REGION Network 43: Barcode - System 3
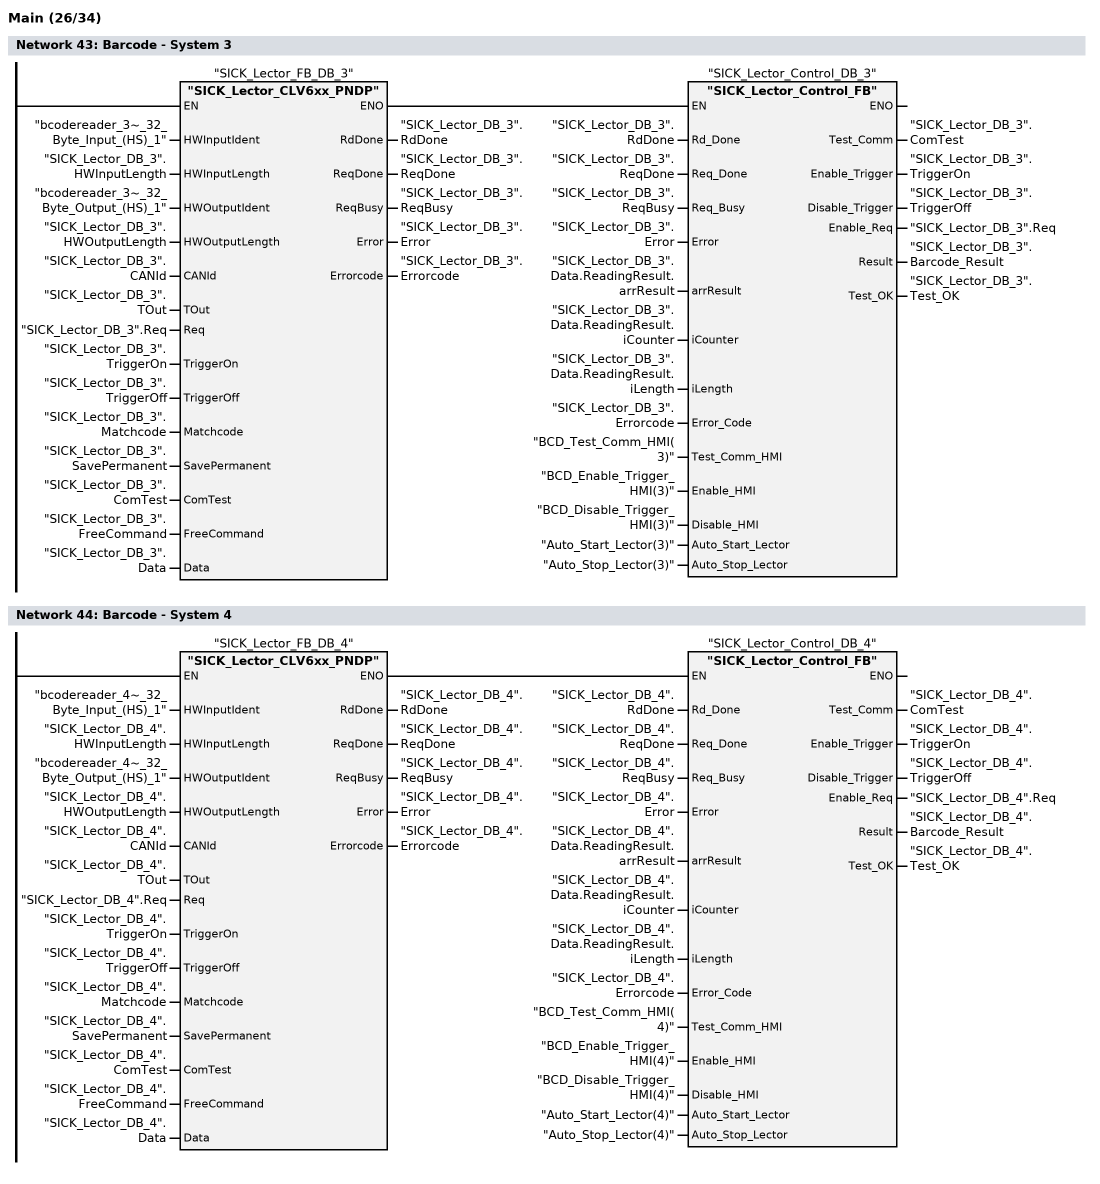
   RUNG wire#powerrail
      "SICK_Lector_FB_DB_3"(HWInputIdent := "bcodereader_3~_32_Byte_Input_(HS)_1", HWInputLength := "SICK_Lector_DB_3".HWInputLength, HWOutputIdent := "bcodereader_3~_32_Byte_Output_(HS)_1", HWOutputLength := "SICK_Lector_DB_3".HWOutputLength, CANId := "SICK_Lector_DB_3".CANId, TOut := "SICK_Lector_DB_3".TOut, Req := "SICK_Lector_DB_3".Req, TriggerOn := "SICK_Lector_DB_3".TriggerOn, TriggerOff := "SICK_Lector_DB_3".TriggerOff, Matchcode := "SICK_Lector_DB_3".Matchcode, SavePermanent := "SICK_Lector_DB_3".SavePermanent, ComTest := "SICK_Lector_DB_3".ComTest, FreeCommand := "SICK_Lector_DB_3".FreeCommand, Data := "SICK_Lector_DB_3".Data, RdDone => "SICK_Lector_DB_3".RdDone, ReqDone => "SICK_Lector_DB_3".ReqDone, ReqBusy => "SICK_Lector_DB_3".ReqBusy, Error => "SICK_Lector_DB_3".Error, Errorcode => "SICK_Lector_DB_3".Errorcode)
      "SICK_Lector_Control_DB_3"(Rd_Done := "SICK_Lector_DB_3".RdDone, Req_Done := "SICK_Lector_DB_3".ReqDone, Req_Busy := "SICK_Lector_DB_3".ReqBusy, Error := "SICK_Lector_DB_3".Error, arrResult := "SICK_Lector_DB_3".Data.ReadingResult.arrResult, iCounter := "SICK_Lector_DB_3".Data.ReadingResult.iCounter, iLength := "SICK_Lector_DB_3".Data.ReadingResult.iLength, Error_Code := "SICK_Lector_DB_3".Errorcode, Test_Comm_HMI := "BCD_Test_Comm_HMI(3)", Enable_HMI := "BCD_Enable_Trigger_HMI(3)", Disable_HMI := "BCD_Disable_Trigger_HMI(3)", Auto_Start_Lector := "Auto_Start_Lector(3)", Auto_Stop_Lector := "Auto_Stop_Lector(3)", Test_Comm => "SICK_Lector_DB_3".ComTest, Enable_Trigger => "SICK_Lector_DB_3".TriggerOn, Disable_Trigger => "SICK_Lector_DB_3".TriggerOff, Enable_Req => "SICK_Lector_DB_3".Req, Result => "SICK_Lector_DB_3".Barcode_Result, Test_OK => "SICK_Lector_DB_3".Test_OK)
   END_RUNG
   // the same network as SCL:
   "SICK_Lector_FB_DB_3"(HWInputIdent := "bcodereader_3~_32_Byte_Input_(HS)_1",   // "SICK_Lector_CLV6xx_PNDP"
                         HWInputLength := "SICK_Lector_DB_3".HWInputLength,
                         HWOutputIdent := "bcodereader_3~_32_Byte_Output_(HS)_1",
                         HWOutputLength := "SICK_Lector_DB_3".HWOutputLength,
                         CANId := "SICK_Lector_DB_3".CANId,
                         TOut := "SICK_Lector_DB_3".TOut,
                         Req := "SICK_Lector_DB_3".Req,
                         TriggerOn := "SICK_Lector_DB_3".TriggerOn,
                         TriggerOff := "SICK_Lector_DB_3".TriggerOff,
                         Matchcode := "SICK_Lector_DB_3".Matchcode,
                         SavePermanent := "SICK_Lector_DB_3".SavePermanent,
                         ComTest := "SICK_Lector_DB_3".ComTest,
                         FreeCommand := "SICK_Lector_DB_3".FreeCommand,
                         Data := "SICK_Lector_DB_3".Data,
                         RdDone => "SICK_Lector_DB_3".RdDone,
                         ReqDone => "SICK_Lector_DB_3".ReqDone,
                         ReqBusy => "SICK_Lector_DB_3".ReqBusy,
                         Error => "SICK_Lector_DB_3".Error,
                         Errorcode => "SICK_Lector_DB_3".Errorcode,
                         ENO => #_w1);
   IF #_w1 THEN
       "SICK_Lector_Control_DB_3"(Rd_Done := "SICK_Lector_DB_3".RdDone,   // "SICK_Lector_Control_FB"
                               Req_Done := "SICK_Lector_DB_3".ReqDone,
                               Req_Busy := "SICK_Lector_DB_3".ReqBusy,
                               Error := "SICK_Lector_DB_3".Error,
                               arrResult := "SICK_Lector_DB_3".Data.ReadingResult.arrResult,
                               iCounter := "SICK_Lector_DB_3".Data.ReadingResult.iCounter,
                               iLength := "SICK_Lector_DB_3".Data.ReadingResult.iLength,
                               Error_Code := "SICK_Lector_DB_3".Errorcode,
                               Test_Comm_HMI := "BCD_Test_Comm_HMI(3)",
                               Enable_HMI := "BCD_Enable_Trigger_HMI(3)",
                               Disable_HMI := "BCD_Disable_Trigger_HMI(3)",
                               Auto_Start_Lector := "Auto_Start_Lector(3)",
                               Auto_Stop_Lector := "Auto_Stop_Lector(3)",
                               Test_Comm => "SICK_Lector_DB_3".ComTest,
                               Enable_Trigger => "SICK_Lector_DB_3".TriggerOn,
                               Disable_Trigger => "SICK_Lector_DB_3".TriggerOff,
                               Enable_Req => "SICK_Lector_DB_3".Req,
                               Result => "SICK_Lector_DB_3".Barcode_Result,
                               Test_OK => "SICK_Lector_DB_3".Test_OK);
   END_IF;
END_REGION

REGION Network 44: Barcode - System 4
   RUNG wire#powerrail
      "SICK_Lector_FB_DB_4"(HWInputIdent := "bcodereader_4~_32_Byte_Input_(HS)_1", HWInputLength := "SICK_Lector_DB_4".HWInputLength, HWOutputIdent := "bcodereader_4~_32_Byte_Output_(HS)_1", HWOutputLength := "SICK_Lector_DB_4".HWOutputLength, CANId := "SICK_Lector_DB_4".CANId, TOut := "SICK_Lector_DB_4".TOut, Req := "SICK_Lector_DB_4".Req, TriggerOn := "SICK_Lector_DB_4".TriggerOn, TriggerOff := "SICK_Lector_DB_4".TriggerOff, Matchcode := "SICK_Lector_DB_4".Matchcode, SavePermanent := "SICK_Lector_DB_4".SavePermanent, ComTest := "SICK_Lector_DB_4".ComTest, FreeCommand := "SICK_Lector_DB_4".FreeCommand, Data := "SICK_Lector_DB_4".Data, RdDone => "SICK_Lector_DB_4".RdDone, ReqDone => "SICK_Lector_DB_4".ReqDone, ReqBusy => "SICK_Lector_DB_4".ReqBusy, Error => "SICK_Lector_DB_4".Error, Errorcode => "SICK_Lector_DB_4".Errorcode)
      "SICK_Lector_Control_DB_4"(Rd_Done := "SICK_Lector_DB_4".RdDone, Req_Done := "SICK_Lector_DB_4".ReqDone, Req_Busy := "SICK_Lector_DB_4".ReqBusy, Error := "SICK_Lector_DB_4".Error, arrResult := "SICK_Lector_DB_4".Data.ReadingResult.arrResult, iCounter := "SICK_Lector_DB_4".Data.ReadingResult.iCounter, iLength := "SICK_Lector_DB_4".Data.ReadingResult.iLength, Error_Code := "SICK_Lector_DB_4".Errorcode, Test_Comm_HMI := "BCD_Test_Comm_HMI(4)", Enable_HMI := "BCD_Enable_Trigger_HMI(4)", Disable_HMI := "BCD_Disable_Trigger_HMI(4)", Auto_Start_Lector := "Auto_Start_Lector(4)", Auto_Stop_Lector := "Auto_Stop_Lector(4)", Test_Comm => "SICK_Lector_DB_4".ComTest, Enable_Trigger => "SICK_Lector_DB_4".TriggerOn, Disable_Trigger => "SICK_Lector_DB_4".TriggerOff, Enable_Req => "SICK_Lector_DB_4".Req, Result => "SICK_Lector_DB_4".Barcode_Result, Test_OK => "SICK_Lector_DB_4".Test_OK)
   END_RUNG
   // the same network as SCL:
   "SICK_Lector_FB_DB_4"(HWInputIdent := "bcodereader_4~_32_Byte_Input_(HS)_1",   // "SICK_Lector_CLV6xx_PNDP"
                         HWInputLength := "SICK_Lector_DB_4".HWInputLength,
                         HWOutputIdent := "bcodereader_4~_32_Byte_Output_(HS)_1",
                         HWOutputLength := "SICK_Lector_DB_4".HWOutputLength,
                         CANId := "SICK_Lector_DB_4".CANId,
                         TOut := "SICK_Lector_DB_4".TOut,
                         Req := "SICK_Lector_DB_4".Req,
                         TriggerOn := "SICK_Lector_DB_4".TriggerOn,
                         TriggerOff := "SICK_Lector_DB_4".TriggerOff,
                         Matchcode := "SICK_Lector_DB_4".Matchcode,
                         SavePermanent := "SICK_Lector_DB_4".SavePermanent,
                         ComTest := "SICK_Lector_DB_4".ComTest,
                         FreeCommand := "SICK_Lector_DB_4".FreeCommand,
                         Data := "SICK_Lector_DB_4".Data,
                         RdDone => "SICK_Lector_DB_4".RdDone,
                         ReqDone => "SICK_Lector_DB_4".ReqDone,
                         ReqBusy => "SICK_Lector_DB_4".ReqBusy,
                         Error => "SICK_Lector_DB_4".Error,
                         Errorcode => "SICK_Lector_DB_4".Errorcode,
                         ENO => #_w1);
   IF #_w1 THEN
       "SICK_Lector_Control_DB_4"(Rd_Done := "SICK_Lector_DB_4".RdDone,   // "SICK_Lector_Control_FB"
                               Req_Done := "SICK_Lector_DB_4".ReqDone,
                               Req_Busy := "SICK_Lector_DB_4".ReqBusy,
                               Error := "SICK_Lector_DB_4".Error,
                               arrResult := "SICK_Lector_DB_4".Data.ReadingResult.arrResult,
                               iCounter := "SICK_Lector_DB_4".Data.ReadingResult.iCounter,
                               iLength := "SICK_Lector_DB_4".Data.ReadingResult.iLength,
                               Error_Code := "SICK_Lector_DB_4".Errorcode,
                               Test_Comm_HMI := "BCD_Test_Comm_HMI(4)",
                               Enable_HMI := "BCD_Enable_Trigger_HMI(4)",
                               Disable_HMI := "BCD_Disable_Trigger_HMI(4)",
                               Auto_Start_Lector := "Auto_Start_Lector(4)",
                               Auto_Stop_Lector := "Auto_Stop_Lector(4)",
                               Test_Comm => "SICK_Lector_DB_4".ComTest,
                               Enable_Trigger => "SICK_Lector_DB_4".TriggerOn,
                               Disable_Trigger => "SICK_Lector_DB_4".TriggerOff,
                               Enable_Req => "SICK_Lector_DB_4".Req,
                               Result => "SICK_Lector_DB_4".Barcode_Result,
                               Test_OK => "SICK_Lector_DB_4".Test_OK);
   END_IF;
END_REGION

REGION Network 45: Barcode - System 5
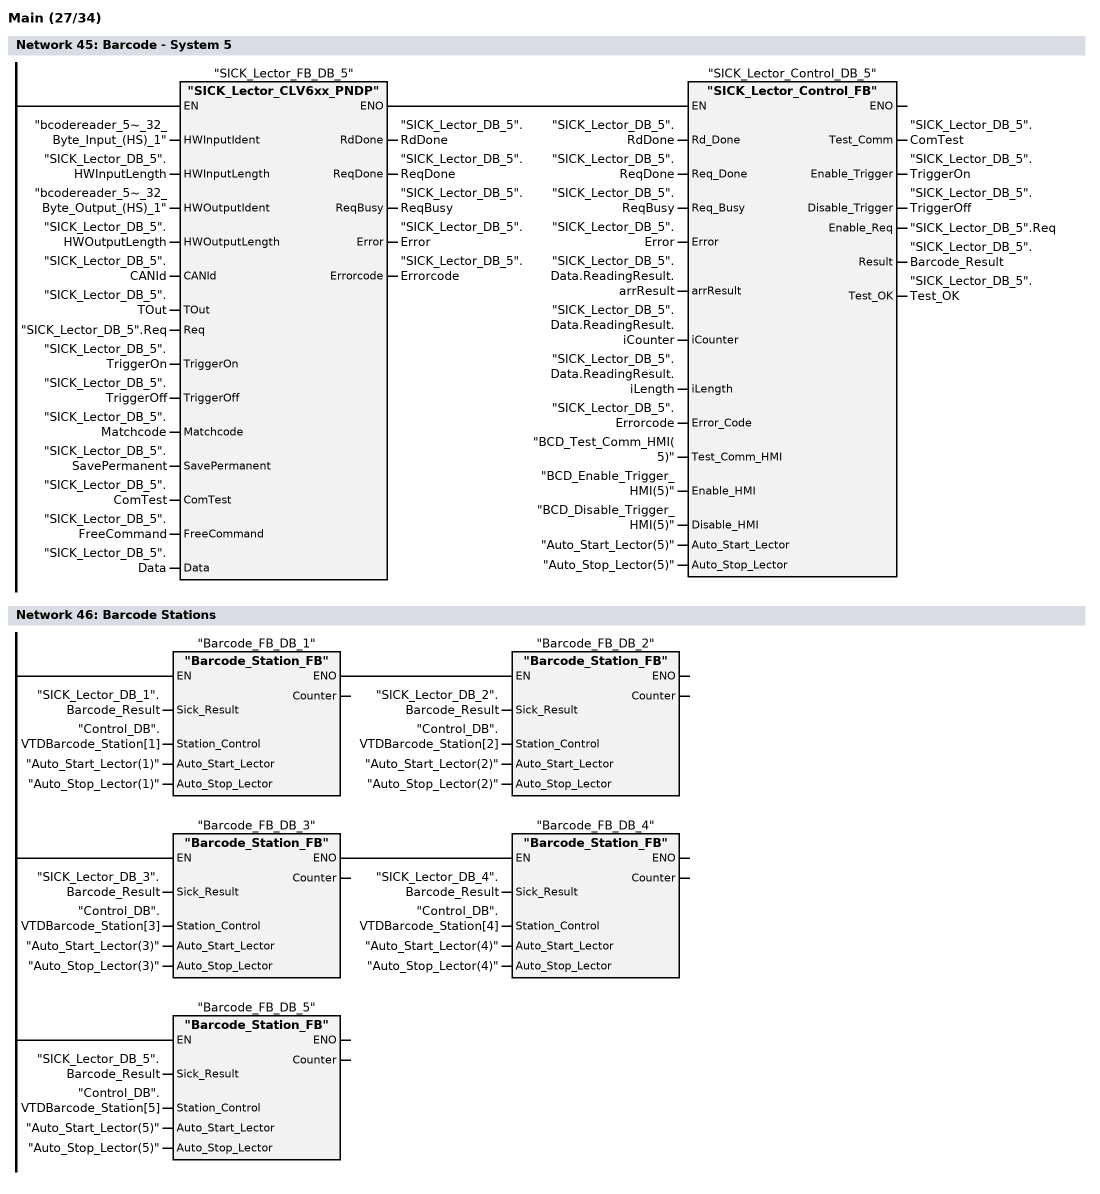
   RUNG wire#powerrail
      "SICK_Lector_FB_DB_5"(HWInputIdent := "bcodereader_5~_32_Byte_Input_(HS)_1", HWInputLength := "SICK_Lector_DB_5".HWInputLength, HWOutputIdent := "bcodereader_5~_32_Byte_Output_(HS)_1", HWOutputLength := "SICK_Lector_DB_5".HWOutputLength, CANId := "SICK_Lector_DB_5".CANId, TOut := "SICK_Lector_DB_5".TOut, Req := "SICK_Lector_DB_5".Req, TriggerOn := "SICK_Lector_DB_5".TriggerOn, TriggerOff := "SICK_Lector_DB_5".TriggerOff, Matchcode := "SICK_Lector_DB_5".Matchcode, SavePermanent := "SICK_Lector_DB_5".SavePermanent, ComTest := "SICK_Lector_DB_5".ComTest, FreeCommand := "SICK_Lector_DB_5".FreeCommand, Data := "SICK_Lector_DB_5".Data, RdDone => "SICK_Lector_DB_5".RdDone, ReqDone => "SICK_Lector_DB_5".ReqDone, ReqBusy => "SICK_Lector_DB_5".ReqBusy, Error => "SICK_Lector_DB_5".Error, Errorcode => "SICK_Lector_DB_5".Errorcode)
      "SICK_Lector_Control_DB_5"(Rd_Done := "SICK_Lector_DB_5".RdDone, Req_Done := "SICK_Lector_DB_5".ReqDone, Req_Busy := "SICK_Lector_DB_5".ReqBusy, Error := "SICK_Lector_DB_5".Error, arrResult := "SICK_Lector_DB_5".Data.ReadingResult.arrResult, iCounter := "SICK_Lector_DB_5".Data.ReadingResult.iCounter, iLength := "SICK_Lector_DB_5".Data.ReadingResult.iLength, Error_Code := "SICK_Lector_DB_5".Errorcode, Test_Comm_HMI := "BCD_Test_Comm_HMI(5)", Enable_HMI := "BCD_Enable_Trigger_HMI(5)", Disable_HMI := "BCD_Disable_Trigger_HMI(5)", Auto_Start_Lector := "Auto_Start_Lector(5)", Auto_Stop_Lector := "Auto_Stop_Lector(5)", Test_Comm => "SICK_Lector_DB_5".ComTest, Enable_Trigger => "SICK_Lector_DB_5".TriggerOn, Disable_Trigger => "SICK_Lector_DB_5".TriggerOff, Enable_Req => "SICK_Lector_DB_5".Req, Result => "SICK_Lector_DB_5".Barcode_Result, Test_OK => "SICK_Lector_DB_5".Test_OK)
   END_RUNG
   // the same network as SCL:
   "SICK_Lector_FB_DB_5"(HWInputIdent := "bcodereader_5~_32_Byte_Input_(HS)_1",   // "SICK_Lector_CLV6xx_PNDP"
                         HWInputLength := "SICK_Lector_DB_5".HWInputLength,
                         HWOutputIdent := "bcodereader_5~_32_Byte_Output_(HS)_1",
                         HWOutputLength := "SICK_Lector_DB_5".HWOutputLength,
                         CANId := "SICK_Lector_DB_5".CANId,
                         TOut := "SICK_Lector_DB_5".TOut,
                         Req := "SICK_Lector_DB_5".Req,
                         TriggerOn := "SICK_Lector_DB_5".TriggerOn,
                         TriggerOff := "SICK_Lector_DB_5".TriggerOff,
                         Matchcode := "SICK_Lector_DB_5".Matchcode,
                         SavePermanent := "SICK_Lector_DB_5".SavePermanent,
                         ComTest := "SICK_Lector_DB_5".ComTest,
                         FreeCommand := "SICK_Lector_DB_5".FreeCommand,
                         Data := "SICK_Lector_DB_5".Data,
                         RdDone => "SICK_Lector_DB_5".RdDone,
                         ReqDone => "SICK_Lector_DB_5".ReqDone,
                         ReqBusy => "SICK_Lector_DB_5".ReqBusy,
                         Error => "SICK_Lector_DB_5".Error,
                         Errorcode => "SICK_Lector_DB_5".Errorcode,
                         ENO => #_w1);
   IF #_w1 THEN
       "SICK_Lector_Control_DB_5"(Rd_Done := "SICK_Lector_DB_5".RdDone,   // "SICK_Lector_Control_FB"
                               Req_Done := "SICK_Lector_DB_5".ReqDone,
                               Req_Busy := "SICK_Lector_DB_5".ReqBusy,
                               Error := "SICK_Lector_DB_5".Error,
                               arrResult := "SICK_Lector_DB_5".Data.ReadingResult.arrResult,
                               iCounter := "SICK_Lector_DB_5".Data.ReadingResult.iCounter,
                               iLength := "SICK_Lector_DB_5".Data.ReadingResult.iLength,
                               Error_Code := "SICK_Lector_DB_5".Errorcode,
                               Test_Comm_HMI := "BCD_Test_Comm_HMI(5)",
                               Enable_HMI := "BCD_Enable_Trigger_HMI(5)",
                               Disable_HMI := "BCD_Disable_Trigger_HMI(5)",
                               Auto_Start_Lector := "Auto_Start_Lector(5)",
                               Auto_Stop_Lector := "Auto_Stop_Lector(5)",
                               Test_Comm => "SICK_Lector_DB_5".ComTest,
                               Enable_Trigger => "SICK_Lector_DB_5".TriggerOn,
                               Disable_Trigger => "SICK_Lector_DB_5".TriggerOff,
                               Enable_Req => "SICK_Lector_DB_5".Req,
                               Result => "SICK_Lector_DB_5".Barcode_Result,
                               Test_OK => "SICK_Lector_DB_5".Test_OK);
   END_IF;
END_REGION

REGION Network 46: Barcode Stations
   RUNG wire#powerrail
      "Barcode_FB_DB_1"(Sick_Result := "SICK_Lector_DB_1".Barcode_Result, Station_Control := "Control_DB".VTDBarcode_Station[1], Auto_Start_Lector := "Auto_Start_Lector(1)", Auto_Stop_Lector := "Auto_Stop_Lector(1)", "Counter" =>)
      "Barcode_FB_DB_2"(Sick_Result := "SICK_Lector_DB_2".Barcode_Result, Station_Control := "Control_DB".VTDBarcode_Station[2], Auto_Start_Lector := "Auto_Start_Lector(2)", Auto_Stop_Lector := "Auto_Stop_Lector(2)", "Counter" =>)
   END_RUNG
   RUNG wire#powerrail
      "Barcode_FB_DB_3"(Sick_Result := "SICK_Lector_DB_3".Barcode_Result, Station_Control := "Control_DB".VTDBarcode_Station[3], Auto_Start_Lector := "Auto_Start_Lector(3)", Auto_Stop_Lector := "Auto_Stop_Lector(3)", "Counter" =>)
      "Barcode_FB_DB_4"(Sick_Result := "SICK_Lector_DB_4".Barcode_Result, Station_Control := "Control_DB".VTDBarcode_Station[4], Auto_Start_Lector := "Auto_Start_Lector(4)", Auto_Stop_Lector := "Auto_Stop_Lector(4)", "Counter" =>)
   END_RUNG
   RUNG wire#powerrail
      "Barcode_FB_DB_5"(Sick_Result := "SICK_Lector_DB_5".Barcode_Result, Station_Control := "Control_DB".VTDBarcode_Station[5], Auto_Start_Lector := "Auto_Start_Lector(5)", Auto_Stop_Lector := "Auto_Stop_Lector(5)", "Counter" =>)
   END_RUNG
   // the same network as SCL:
   "Barcode_FB_DB_1"(Sick_Result := "SICK_Lector_DB_1".Barcode_Result,   // "Barcode_Station_FB"
                     Station_Control := "Control_DB".VTDBarcode_Station[1],
                     Auto_Start_Lector := "Auto_Start_Lector(1)",
                     Auto_Stop_Lector := "Auto_Stop_Lector(1)",
                     ENO => #_w1);
   IF #_w1 THEN
       "Barcode_FB_DB_2"(Sick_Result := "SICK_Lector_DB_2".Barcode_Result,   // "Barcode_Station_FB"
                         Station_Control := "Control_DB".VTDBarcode_Station[2],
                         Auto_Start_Lector := "Auto_Start_Lector(2)",
                         Auto_Stop_Lector := "Auto_Stop_Lector(2)");
   END_IF;
   "Barcode_FB_DB_3"(Sick_Result := "SICK_Lector_DB_3".Barcode_Result,   // "Barcode_Station_FB"
                     Station_Control := "Control_DB".VTDBarcode_Station[3],
                     Auto_Start_Lector := "Auto_Start_Lector(3)",
                     Auto_Stop_Lector := "Auto_Stop_Lector(3)",
                     ENO => #_w2);
   IF #_w2 THEN
       "Barcode_FB_DB_4"(Sick_Result := "SICK_Lector_DB_4".Barcode_Result,   // "Barcode_Station_FB"
                         Station_Control := "Control_DB".VTDBarcode_Station[4],
                         Auto_Start_Lector := "Auto_Start_Lector(4)",
                         Auto_Stop_Lector := "Auto_Stop_Lector(4)");
   END_IF;
   "Barcode_FB_DB_5"(Sick_Result := "SICK_Lector_DB_5".Barcode_Result,   // "Barcode_Station_FB"
                     Station_Control := "Control_DB".VTDBarcode_Station[5],
                     Auto_Start_Lector := "Auto_Start_Lector(5)",
                     Auto_Stop_Lector := "Auto_Stop_Lector(5)");
END_REGION

REGION Network 47: Stack Lights
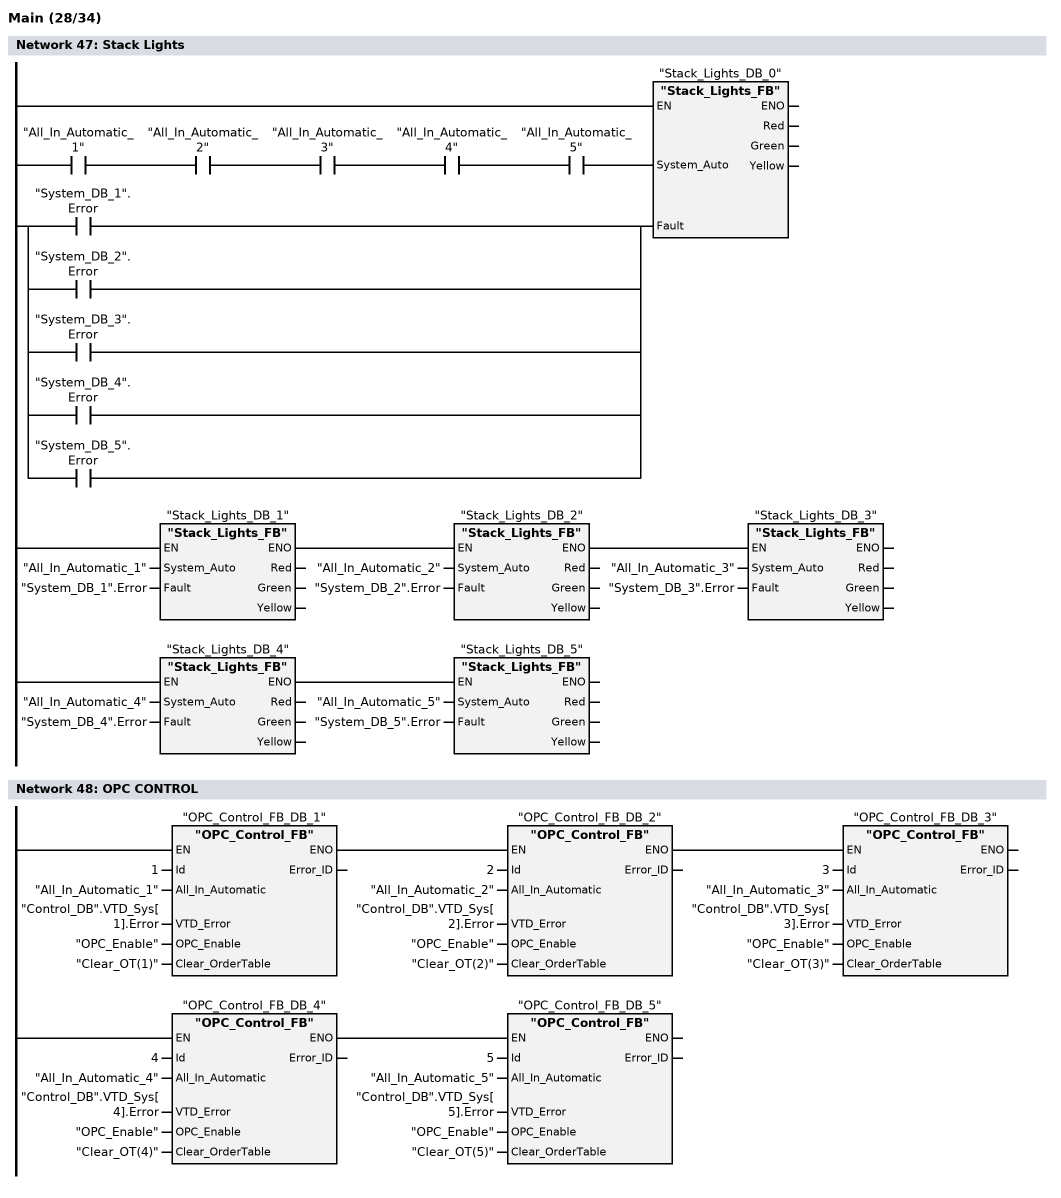
   RUNG wire#powerrail
      "Stack_Lights_DB_0"(System_Auto := wire#w1, Fault := wire#w2, Red =>, Green =>, Yellow =>)
   END_RUNG
   RUNG wire#powerrail
      Contact( "All_In_Automatic_1" )
      Contact( "All_In_Automatic_2" )
      Contact( "All_In_Automatic_3" )
      Contact( "All_In_Automatic_4" )
      Contact( "All_In_Automatic_5" )
   END_RUNG wire#w1
   RUNG wire#powerrail
      Contact( "System_DB_1".Error )
   END_RUNG wire#w2
   RUNG wire#powerrail
      Contact( "System_DB_2".Error )
   END_RUNG wire#w2
   RUNG wire#powerrail
      Contact( "System_DB_3".Error )
   END_RUNG wire#w2
   RUNG wire#powerrail
      Contact( "System_DB_4".Error )
   END_RUNG wire#w2
   RUNG wire#powerrail
      Contact( "System_DB_5".Error )
   END_RUNG wire#w2
   RUNG wire#powerrail
      "Stack_Lights_DB_1"(System_Auto := "All_In_Automatic_1", Fault := "System_DB_1".Error, Red =>, Green =>, Yellow =>)
      "Stack_Lights_DB_2"(System_Auto := "All_In_Automatic_2", Fault := "System_DB_2".Error, Red =>, Green =>, Yellow =>)
      "Stack_Lights_DB_3"(System_Auto := "All_In_Automatic_3", Fault := "System_DB_3".Error, Red =>, Green =>, Yellow =>)
   END_RUNG
   RUNG wire#powerrail
      "Stack_Lights_DB_4"(System_Auto := "All_In_Automatic_4", Fault := "System_DB_4".Error, Red =>, Green =>, Yellow =>)
      "Stack_Lights_DB_5"(System_Auto := "All_In_Automatic_5", Fault := "System_DB_5".Error, Red =>, Green =>, Yellow =>)
   END_RUNG
   // the same network as SCL:
   "Stack_Lights_DB_0"(System_Auto := "All_In_Automatic_1" AND "All_In_Automatic_2" AND "All_In_Automatic_3" AND "All_In_Automatic_4" AND "All_In_Automatic_5",   // "Stack_Lights_FB"
                       Fault := "System_DB_1".Error OR "System_DB_2".Error OR "System_DB_3".Error OR "System_DB_4".Error OR "System_DB_5".Error);
   "Stack_Lights_DB_1"(System_Auto := "All_In_Automatic_1", Fault := "System_DB_1".Error, ENO => #_w1);   // "Stack_Lights_FB"
   "Stack_Lights_DB_2"(EN := #_w1,   // "Stack_Lights_FB"
                       System_Auto := "All_In_Automatic_2",
                       Fault := "System_DB_2".Error,
                       ENO => #_w2);
   IF #_w2 THEN
       "Stack_Lights_DB_3"(System_Auto := "All_In_Automatic_3", Fault := "System_DB_3".Error);   // "Stack_Lights_FB"
   END_IF;
   "Stack_Lights_DB_4"(System_Auto := "All_In_Automatic_4", Fault := "System_DB_4".Error, ENO => #_w3);   // "Stack_Lights_FB"
   IF #_w3 THEN
       "Stack_Lights_DB_5"(System_Auto := "All_In_Automatic_5", Fault := "System_DB_5".Error);   // "Stack_Lights_FB"
   END_IF;
END_REGION

REGION Network 48: OPC CONTROL
   RUNG wire#powerrail
      "OPC_Control_FB_DB_1"(Id := 1, All_In_Automatic := "All_In_Automatic_1", VTD_Error := "Control_DB".VTD_Sys[1].Error, OPC_Enable := "OPC_Enable", Clear_OrderTable := "Clear_OT(1)", Error_ID =>)
      "OPC_Control_FB_DB_2"(Id := 2, All_In_Automatic := "All_In_Automatic_2", VTD_Error := "Control_DB".VTD_Sys[2].Error, OPC_Enable := "OPC_Enable", Clear_OrderTable := "Clear_OT(2)", Error_ID =>)
      "OPC_Control_FB_DB_3"(Id := 3, All_In_Automatic := "All_In_Automatic_3", VTD_Error := "Control_DB".VTD_Sys[3].Error, OPC_Enable := "OPC_Enable", Clear_OrderTable := "Clear_OT(3)", Error_ID =>)
   END_RUNG
   RUNG wire#powerrail
      "OPC_Control_FB_DB_4"(Id := 4, All_In_Automatic := "All_In_Automatic_4", VTD_Error := "Control_DB".VTD_Sys[4].Error, OPC_Enable := "OPC_Enable", Clear_OrderTable := "Clear_OT(4)", Error_ID =>)
      "OPC_Control_FB_DB_5"(Id := 5, All_In_Automatic := "All_In_Automatic_5", VTD_Error := "Control_DB".VTD_Sys[5].Error, OPC_Enable := "OPC_Enable", Clear_OrderTable := "Clear_OT(5)", Error_ID =>)
   END_RUNG
   // the same network as SCL:
   "OPC_Control_FB_DB_1"(Id := 1,   // "OPC_Control_FB"
                         All_In_Automatic := "All_In_Automatic_1",
                         VTD_Error := "Control_DB".VTD_Sys[1].Error,
                         OPC_Enable := "OPC_Enable",
                         Clear_OrderTable := "Clear_OT(1)",
                         ENO => #_w1);
   "OPC_Control_FB_DB_2"(EN := #_w1,   // "OPC_Control_FB"
                         Id := 2,
                         All_In_Automatic := "All_In_Automatic_2",
                         VTD_Error := "Control_DB".VTD_Sys[2].Error,
                         OPC_Enable := "OPC_Enable",
                         Clear_OrderTable := "Clear_OT(2)",
                         ENO => #_w2);
   IF #_w2 THEN
       "OPC_Control_FB_DB_3"(Id := 3,   // "OPC_Control_FB"
                             All_In_Automatic := "All_In_Automatic_3",
                             VTD_Error := "Control_DB".VTD_Sys[3].Error,
                             OPC_Enable := "OPC_Enable",
                             Clear_OrderTable := "Clear_OT(3)");
   END_IF;
   "OPC_Control_FB_DB_4"(Id := 4,   // "OPC_Control_FB"
                         All_In_Automatic := "All_In_Automatic_4",
                         VTD_Error := "Control_DB".VTD_Sys[4].Error,
                         OPC_Enable := "OPC_Enable",
                         Clear_OrderTable := "Clear_OT(4)",
                         ENO => #_w3);
   IF #_w3 THEN
       "OPC_Control_FB_DB_5"(Id := 5,   // "OPC_Control_FB"
                             All_In_Automatic := "All_In_Automatic_5",
                             VTD_Error := "Control_DB".VTD_Sys[5].Error,
                             OPC_Enable := "OPC_Enable",
                             Clear_OrderTable := "Clear_OT(5)");
   END_IF;
END_REGION

REGION Network 49: Shuttle TCPs
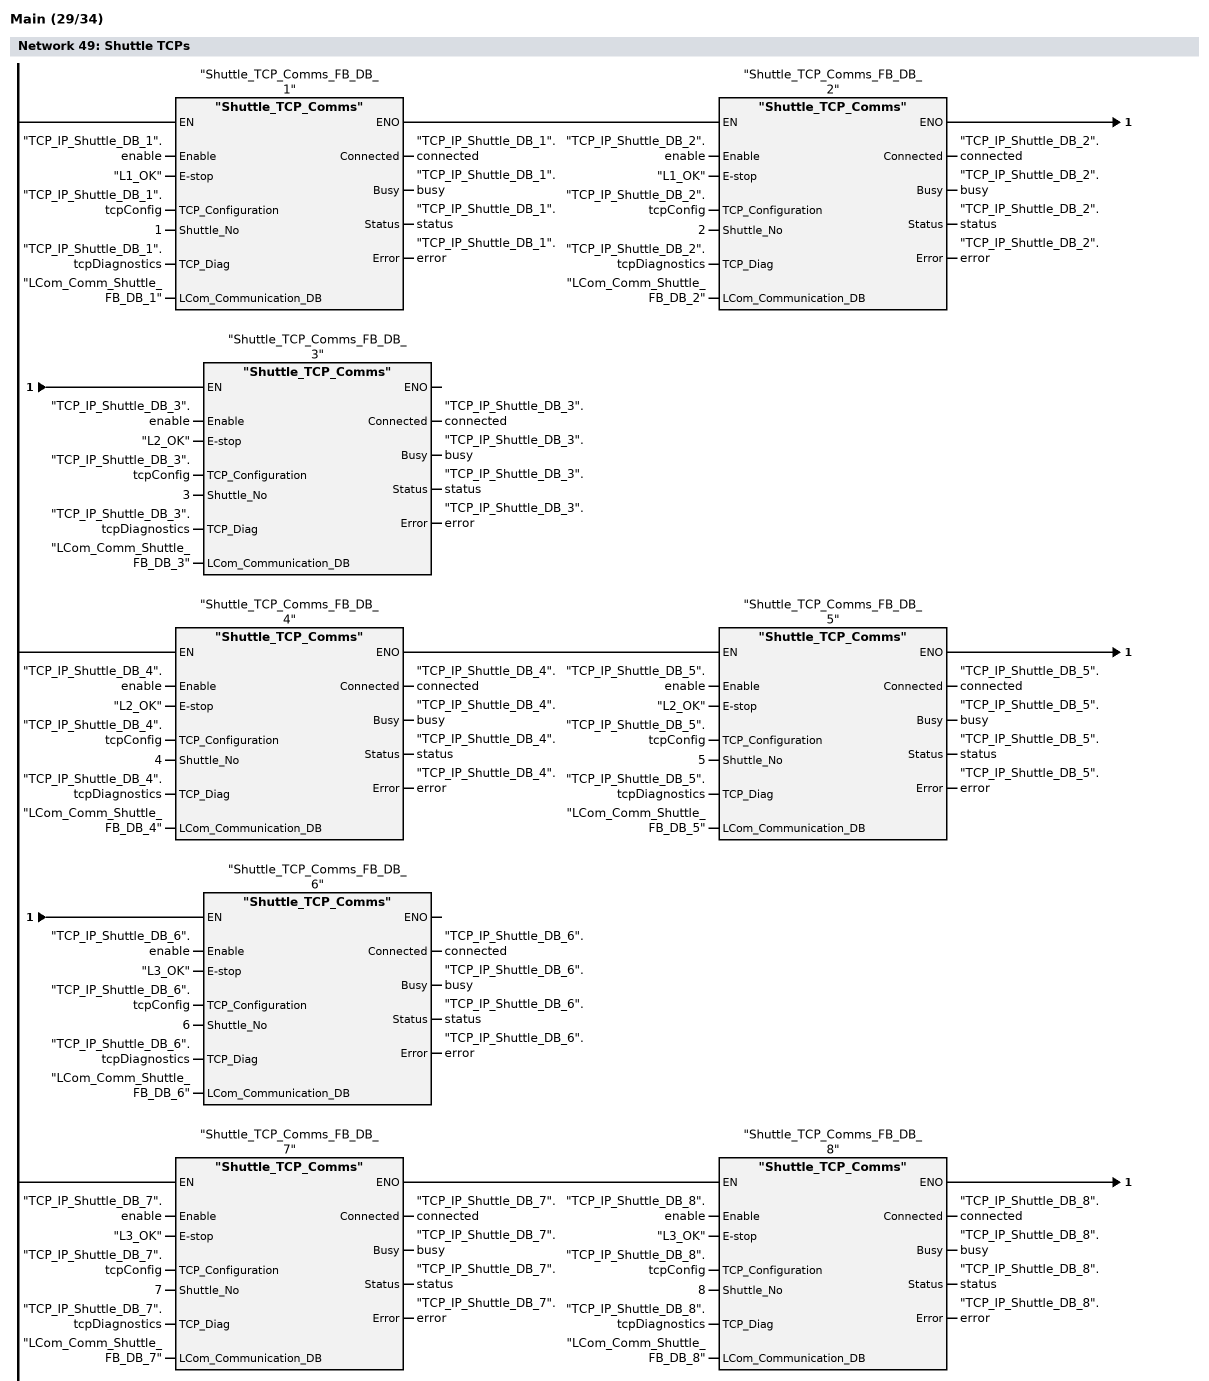
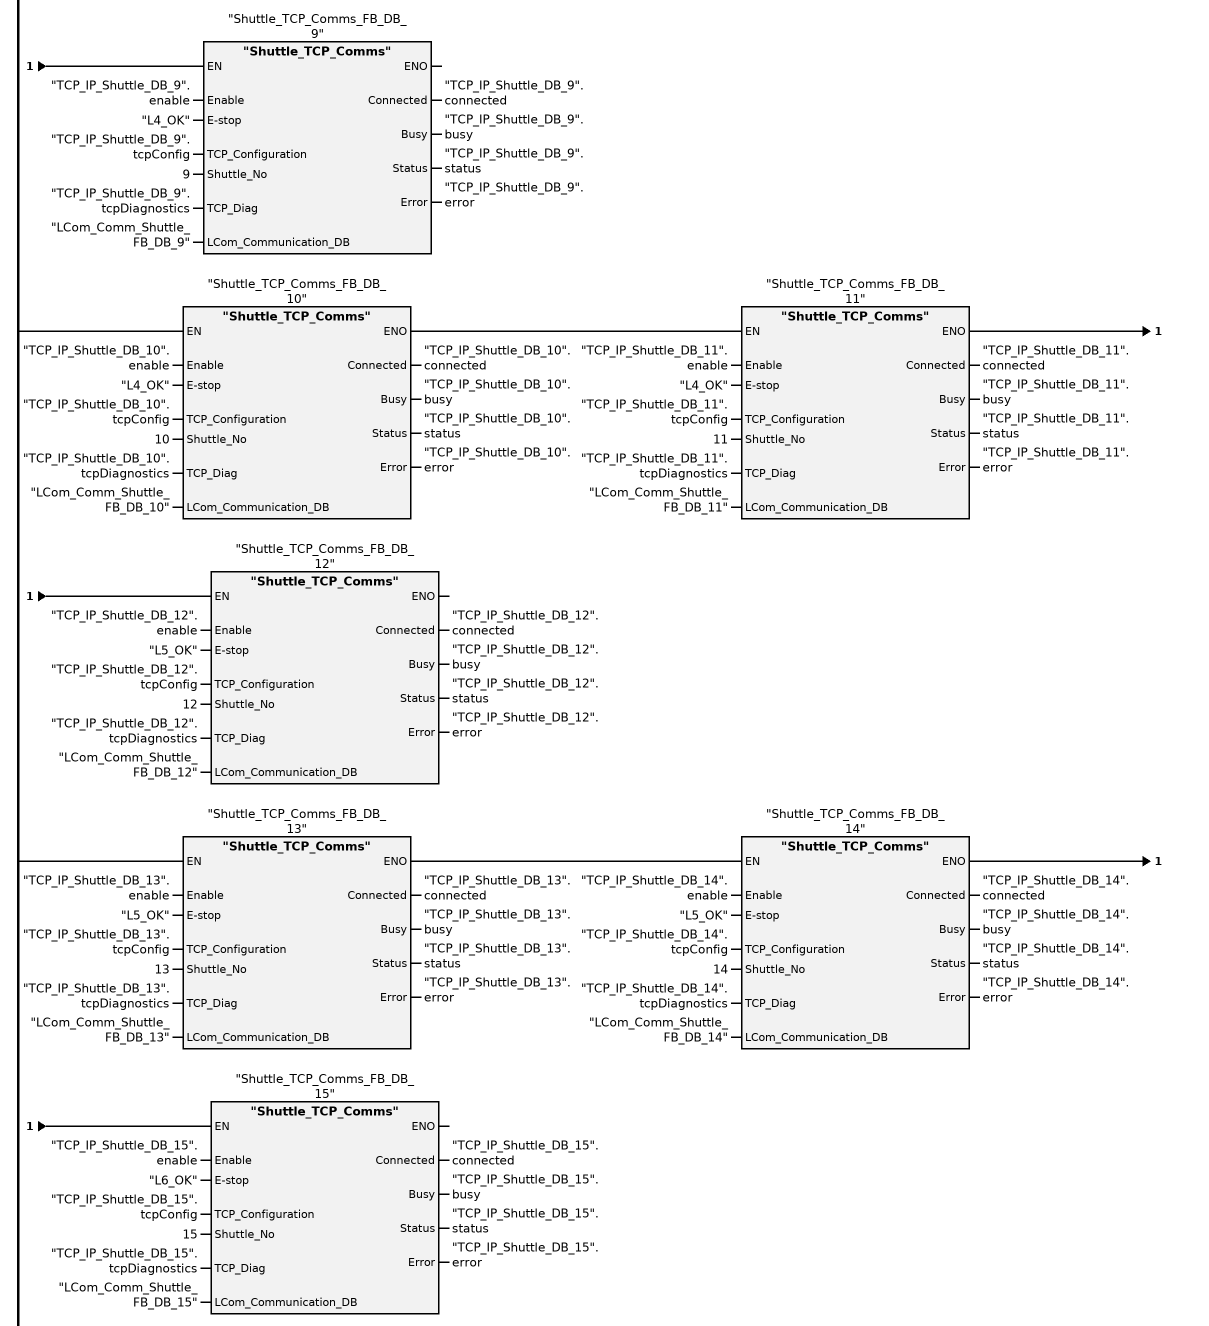
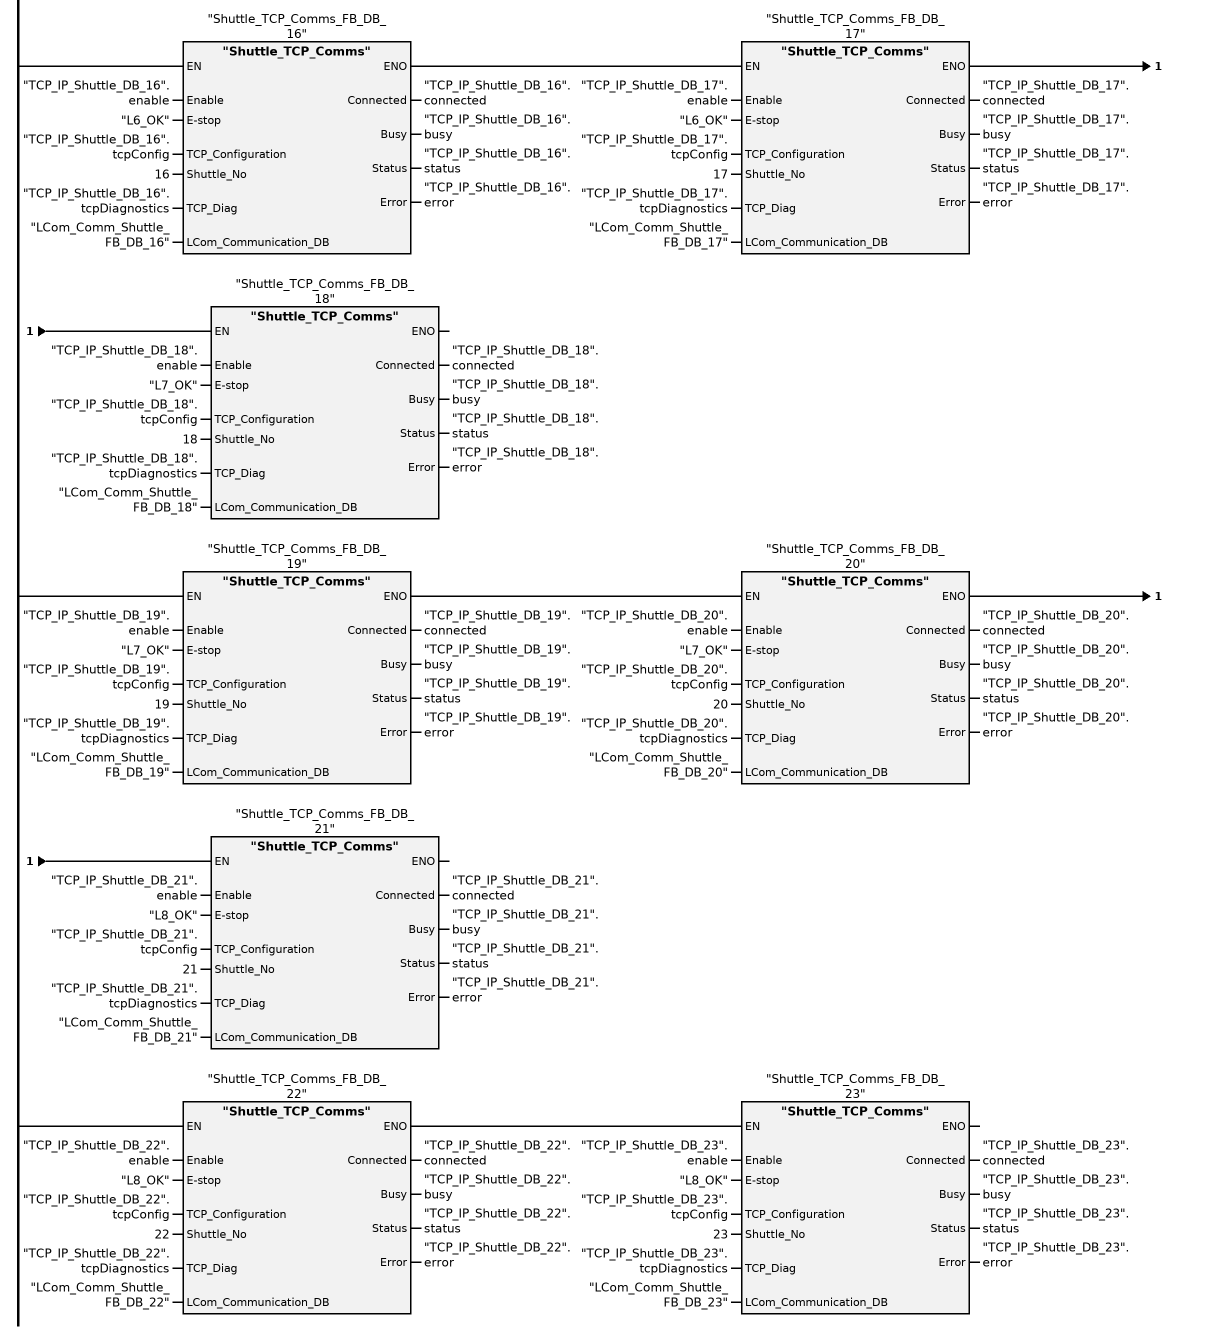
   RUNG wire#powerrail
      "Shuttle_TCP_Comms_FB_DB_1"(Enable := "TCP_IP_Shuttle_DB_1".enable, "E-stop" := "L1_OK", TCP_Configuration := "TCP_IP_Shuttle_DB_1".tcpConfig, Shuttle_No := 1, TCP_Diag := "TCP_IP_Shuttle_DB_1".tcpDiagnostics, LCom_Communication_DB := "LCom_Comm_Shuttle_FB_DB_1", Connected => "TCP_IP_Shuttle_DB_1".connected, Busy => "TCP_IP_Shuttle_DB_1".busy, Status => "TCP_IP_Shuttle_DB_1".status, Error => "TCP_IP_Shuttle_DB_1".error)
      "Shuttle_TCP_Comms_FB_DB_2"(Enable := "TCP_IP_Shuttle_DB_2".enable, "E-stop" := "L1_OK", TCP_Configuration := "TCP_IP_Shuttle_DB_2".tcpConfig, Shuttle_No := 2, TCP_Diag := "TCP_IP_Shuttle_DB_2".tcpDiagnostics, LCom_Communication_DB := "LCom_Comm_Shuttle_FB_DB_2", Connected => "TCP_IP_Shuttle_DB_2".connected, Busy => "TCP_IP_Shuttle_DB_2".busy, Status => "TCP_IP_Shuttle_DB_2".status, Error => "TCP_IP_Shuttle_DB_2".error)
      "Shuttle_TCP_Comms_FB_DB_3"(Enable := "TCP_IP_Shuttle_DB_3".enable, "E-stop" := "L2_OK", TCP_Configuration := "TCP_IP_Shuttle_DB_3".tcpConfig, Shuttle_No := 3, TCP_Diag := "TCP_IP_Shuttle_DB_3".tcpDiagnostics, LCom_Communication_DB := "LCom_Comm_Shuttle_FB_DB_3", Connected => "TCP_IP_Shuttle_DB_3".connected, Busy => "TCP_IP_Shuttle_DB_3".busy, Status => "TCP_IP_Shuttle_DB_3".status, Error => "TCP_IP_Shuttle_DB_3".error)
   END_RUNG
   RUNG wire#powerrail
      "Shuttle_TCP_Comms_FB_DB_4"(Enable := "TCP_IP_Shuttle_DB_4".enable, "E-stop" := "L2_OK", TCP_Configuration := "TCP_IP_Shuttle_DB_4".tcpConfig, Shuttle_No := 4, TCP_Diag := "TCP_IP_Shuttle_DB_4".tcpDiagnostics, LCom_Communication_DB := "LCom_Comm_Shuttle_FB_DB_4", Connected => "TCP_IP_Shuttle_DB_4".connected, Busy => "TCP_IP_Shuttle_DB_4".busy, Status => "TCP_IP_Shuttle_DB_4".status, Error => "TCP_IP_Shuttle_DB_4".error)
      "Shuttle_TCP_Comms_FB_DB_5"(Enable := "TCP_IP_Shuttle_DB_5".enable, "E-stop" := "L2_OK", TCP_Configuration := "TCP_IP_Shuttle_DB_5".tcpConfig, Shuttle_No := 5, TCP_Diag := "TCP_IP_Shuttle_DB_5".tcpDiagnostics, LCom_Communication_DB := "LCom_Comm_Shuttle_FB_DB_5", Connected => "TCP_IP_Shuttle_DB_5".connected, Busy => "TCP_IP_Shuttle_DB_5".busy, Status => "TCP_IP_Shuttle_DB_5".status, Error => "TCP_IP_Shuttle_DB_5".error)
      "Shuttle_TCP_Comms_FB_DB_6"(Enable := "TCP_IP_Shuttle_DB_6".enable, "E-stop" := "L3_OK", TCP_Configuration := "TCP_IP_Shuttle_DB_6".tcpConfig, Shuttle_No := 6, TCP_Diag := "TCP_IP_Shuttle_DB_6".tcpDiagnostics, LCom_Communication_DB := "LCom_Comm_Shuttle_FB_DB_6", Connected => "TCP_IP_Shuttle_DB_6".connected, Busy => "TCP_IP_Shuttle_DB_6".busy, Status => "TCP_IP_Shuttle_DB_6".status, Error => "TCP_IP_Shuttle_DB_6".error)
   END_RUNG
   RUNG wire#powerrail
      "Shuttle_TCP_Comms_FB_DB_7"(Enable := "TCP_IP_Shuttle_DB_7".enable, "E-stop" := "L3_OK", TCP_Configuration := "TCP_IP_Shuttle_DB_7".tcpConfig, Shuttle_No := 7, TCP_Diag := "TCP_IP_Shuttle_DB_7".tcpDiagnostics, LCom_Communication_DB := "LCom_Comm_Shuttle_FB_DB_7", Connected => "TCP_IP_Shuttle_DB_7".connected, Busy => "TCP_IP_Shuttle_DB_7".busy, Status => "TCP_IP_Shuttle_DB_7".status, Error => "TCP_IP_Shuttle_DB_7".error)
      "Shuttle_TCP_Comms_FB_DB_8"(Enable := "TCP_IP_Shuttle_DB_8".enable, "E-stop" := "L3_OK", TCP_Configuration := "TCP_IP_Shuttle_DB_8".tcpConfig, Shuttle_No := 8, TCP_Diag := "TCP_IP_Shuttle_DB_8".tcpDiagnostics, LCom_Communication_DB := "LCom_Comm_Shuttle_FB_DB_8", Connected => "TCP_IP_Shuttle_DB_8".connected, Busy => "TCP_IP_Shuttle_DB_8".busy, Status => "TCP_IP_Shuttle_DB_8".status, Error => "TCP_IP_Shuttle_DB_8".error)
      "Shuttle_TCP_Comms_FB_DB_9"(Enable := "TCP_IP_Shuttle_DB_9".enable, "E-stop" := "L4_OK", TCP_Configuration := "TCP_IP_Shuttle_DB_9".tcpConfig, Shuttle_No := 9, TCP_Diag := "TCP_IP_Shuttle_DB_9".tcpDiagnostics, LCom_Communication_DB := "LCom_Comm_Shuttle_FB_DB_9", Connected => "TCP_IP_Shuttle_DB_9".connected, Busy => "TCP_IP_Shuttle_DB_9".busy, Status => "TCP_IP_Shuttle_DB_9".status, Error => "TCP_IP_Shuttle_DB_9".error)
   END_RUNG
   RUNG wire#powerrail
      "Shuttle_TCP_Comms_FB_DB_10"(Enable := "TCP_IP_Shuttle_DB_10".enable, "E-stop" := "L4_OK", TCP_Configuration := "TCP_IP_Shuttle_DB_10".tcpConfig, Shuttle_No := 10, TCP_Diag := "TCP_IP_Shuttle_DB_10".tcpDiagnostics, LCom_Communication_DB := "LCom_Comm_Shuttle_FB_DB_10", Connected => "TCP_IP_Shuttle_DB_10".connected, Busy => "TCP_IP_Shuttle_DB_10".busy, Status => "TCP_IP_Shuttle_DB_10".status, Error => "TCP_IP_Shuttle_DB_10".error)
      "Shuttle_TCP_Comms_FB_DB_11"(Enable := "TCP_IP_Shuttle_DB_11".enable, "E-stop" := "L4_OK", TCP_Configuration := "TCP_IP_Shuttle_DB_11".tcpConfig, Shuttle_No := 11, TCP_Diag := "TCP_IP_Shuttle_DB_11".tcpDiagnostics, LCom_Communication_DB := "LCom_Comm_Shuttle_FB_DB_11", Connected => "TCP_IP_Shuttle_DB_11".connected, Busy => "TCP_IP_Shuttle_DB_11".busy, Status => "TCP_IP_Shuttle_DB_11".status, Error => "TCP_IP_Shuttle_DB_11".error)
      "Shuttle_TCP_Comms_FB_DB_12"(Enable := "TCP_IP_Shuttle_DB_12".enable, "E-stop" := "L5_OK", TCP_Configuration := "TCP_IP_Shuttle_DB_12".tcpConfig, Shuttle_No := 12, TCP_Diag := "TCP_IP_Shuttle_DB_12".tcpDiagnostics, LCom_Communication_DB := "LCom_Comm_Shuttle_FB_DB_12", Connected => "TCP_IP_Shuttle_DB_12".connected, Busy => "TCP_IP_Shuttle_DB_12".busy, Status => "TCP_IP_Shuttle_DB_12".status, Error => "TCP_IP_Shuttle_DB_12".error)
   END_RUNG
   RUNG wire#powerrail
      "Shuttle_TCP_Comms_FB_DB_13"(Enable := "TCP_IP_Shuttle_DB_13".enable, "E-stop" := "L5_OK", TCP_Configuration := "TCP_IP_Shuttle_DB_13".tcpConfig, Shuttle_No := 13, TCP_Diag := "TCP_IP_Shuttle_DB_13".tcpDiagnostics, LCom_Communication_DB := "LCom_Comm_Shuttle_FB_DB_13", Connected => "TCP_IP_Shuttle_DB_13".connected, Busy => "TCP_IP_Shuttle_DB_13".busy, Status => "TCP_IP_Shuttle_DB_13".status, Error => "TCP_IP_Shuttle_DB_13".error)
      "Shuttle_TCP_Comms_FB_DB_14"(Enable := "TCP_IP_Shuttle_DB_14".enable, "E-stop" := "L5_OK", TCP_Configuration := "TCP_IP_Shuttle_DB_14".tcpConfig, Shuttle_No := 14, TCP_Diag := "TCP_IP_Shuttle_DB_14".tcpDiagnostics, LCom_Communication_DB := "LCom_Comm_Shuttle_FB_DB_14", Connected => "TCP_IP_Shuttle_DB_14".connected, Busy => "TCP_IP_Shuttle_DB_14".busy, Status => "TCP_IP_Shuttle_DB_14".status, Error => "TCP_IP_Shuttle_DB_14".error)
      "Shuttle_TCP_Comms_FB_DB_15"(Enable := "TCP_IP_Shuttle_DB_15".enable, "E-stop" := "L6_OK", TCP_Configuration := "TCP_IP_Shuttle_DB_15".tcpConfig, Shuttle_No := 15, TCP_Diag := "TCP_IP_Shuttle_DB_15".tcpDiagnostics, LCom_Communication_DB := "LCom_Comm_Shuttle_FB_DB_15", Connected => "TCP_IP_Shuttle_DB_15".connected, Busy => "TCP_IP_Shuttle_DB_15".busy, Status => "TCP_IP_Shuttle_DB_15".status, Error => "TCP_IP_Shuttle_DB_15".error)
   END_RUNG
   RUNG wire#powerrail
      "Shuttle_TCP_Comms_FB_DB_16"(Enable := "TCP_IP_Shuttle_DB_16".enable, "E-stop" := "L6_OK", TCP_Configuration := "TCP_IP_Shuttle_DB_16".tcpConfig, Shuttle_No := 16, TCP_Diag := "TCP_IP_Shuttle_DB_16".tcpDiagnostics, LCom_Communication_DB := "LCom_Comm_Shuttle_FB_DB_16", Connected => "TCP_IP_Shuttle_DB_16".connected, Busy => "TCP_IP_Shuttle_DB_16".busy, Status => "TCP_IP_Shuttle_DB_16".status, Error => "TCP_IP_Shuttle_DB_16".error)
      "Shuttle_TCP_Comms_FB_DB_17"(Enable := "TCP_IP_Shuttle_DB_17".enable, "E-stop" := "L6_OK", TCP_Configuration := "TCP_IP_Shuttle_DB_17".tcpConfig, Shuttle_No := 17, TCP_Diag := "TCP_IP_Shuttle_DB_17".tcpDiagnostics, LCom_Communication_DB := "LCom_Comm_Shuttle_FB_DB_17", Connected => "TCP_IP_Shuttle_DB_17".connected, Busy => "TCP_IP_Shuttle_DB_17".busy, Status => "TCP_IP_Shuttle_DB_17".status, Error => "TCP_IP_Shuttle_DB_17".error)
      "Shuttle_TCP_Comms_FB_DB_18"(Enable := "TCP_IP_Shuttle_DB_18".enable, "E-stop" := "L7_OK", TCP_Configuration := "TCP_IP_Shuttle_DB_18".tcpConfig, Shuttle_No := 18, TCP_Diag := "TCP_IP_Shuttle_DB_18".tcpDiagnostics, LCom_Communication_DB := "LCom_Comm_Shuttle_FB_DB_18", Connected => "TCP_IP_Shuttle_DB_18".connected, Busy => "TCP_IP_Shuttle_DB_18".busy, Status => "TCP_IP_Shuttle_DB_18".status, Error => "TCP_IP_Shuttle_DB_18".error)
   END_RUNG
   RUNG wire#powerrail
      "Shuttle_TCP_Comms_FB_DB_19"(Enable := "TCP_IP_Shuttle_DB_19".enable, "E-stop" := "L7_OK", TCP_Configuration := "TCP_IP_Shuttle_DB_19".tcpConfig, Shuttle_No := 19, TCP_Diag := "TCP_IP_Shuttle_DB_19".tcpDiagnostics, LCom_Communication_DB := "LCom_Comm_Shuttle_FB_DB_19", Connected => "TCP_IP_Shuttle_DB_19".connected, Busy => "TCP_IP_Shuttle_DB_19".busy, Status => "TCP_IP_Shuttle_DB_19".status, Error => "TCP_IP_Shuttle_DB_19".error)
      "Shuttle_TCP_Comms_FB_DB_20"(Enable := "TCP_IP_Shuttle_DB_20".enable, "E-stop" := "L7_OK", TCP_Configuration := "TCP_IP_Shuttle_DB_20".tcpConfig, Shuttle_No := 20, TCP_Diag := "TCP_IP_Shuttle_DB_20".tcpDiagnostics, LCom_Communication_DB := "LCom_Comm_Shuttle_FB_DB_20", Connected => "TCP_IP_Shuttle_DB_20".connected, Busy => "TCP_IP_Shuttle_DB_20".busy, Status => "TCP_IP_Shuttle_DB_20".status, Error => "TCP_IP_Shuttle_DB_20".error)
      "Shuttle_TCP_Comms_FB_DB_21"(Enable := "TCP_IP_Shuttle_DB_21".enable, "E-stop" := "L8_OK", TCP_Configuration := "TCP_IP_Shuttle_DB_21".tcpConfig, Shuttle_No := 21, TCP_Diag := "TCP_IP_Shuttle_DB_21".tcpDiagnostics, LCom_Communication_DB := "LCom_Comm_Shuttle_FB_DB_21", Connected => "TCP_IP_Shuttle_DB_21".connected, Busy => "TCP_IP_Shuttle_DB_21".busy, Status => "TCP_IP_Shuttle_DB_21".status, Error => "TCP_IP_Shuttle_DB_21".error)
   END_RUNG
   RUNG wire#powerrail
      "Shuttle_TCP_Comms_FB_DB_22"(Enable := "TCP_IP_Shuttle_DB_22".enable, "E-stop" := "L8_OK", TCP_Configuration := "TCP_IP_Shuttle_DB_22".tcpConfig, Shuttle_No := 22, TCP_Diag := "TCP_IP_Shuttle_DB_22".tcpDiagnostics, LCom_Communication_DB := "LCom_Comm_Shuttle_FB_DB_22", Connected => "TCP_IP_Shuttle_DB_22".connected, Busy => "TCP_IP_Shuttle_DB_22".busy, Status => "TCP_IP_Shuttle_DB_22".status, Error => "TCP_IP_Shuttle_DB_22".error)
      "Shuttle_TCP_Comms_FB_DB_23"(Enable := "TCP_IP_Shuttle_DB_23".enable, "E-stop" := "L8_OK", TCP_Configuration := "TCP_IP_Shuttle_DB_23".tcpConfig, Shuttle_No := 23, TCP_Diag := "TCP_IP_Shuttle_DB_23".tcpDiagnostics, LCom_Communication_DB := "LCom_Comm_Shuttle_FB_DB_23", Connected => "TCP_IP_Shuttle_DB_23".connected, Busy => "TCP_IP_Shuttle_DB_23".busy, Status => "TCP_IP_Shuttle_DB_23".status, Error => "TCP_IP_Shuttle_DB_23".error)
   END_RUNG
   // the same network as SCL:
   "Shuttle_TCP_Comms_FB_DB_1"(Enable := "TCP_IP_Shuttle_DB_1".enable,   // "Shuttle_TCP_Comms"
                           "E-stop" := "L1_OK",
                           TCP_Configuration := "TCP_IP_Shuttle_DB_1".tcpConfig,
                           Shuttle_No := 1,
                           TCP_Diag := "TCP_IP_Shuttle_DB_1".tcpDiagnostics,
                           LCom_Communication_DB := "LCom_Comm_Shuttle_FB_DB_1",
                           Connected => "TCP_IP_Shuttle_DB_1".connected,
                           Busy => "TCP_IP_Shuttle_DB_1".busy,
                           Status => "TCP_IP_Shuttle_DB_1".status,
                           Error => "TCP_IP_Shuttle_DB_1".error,
                           ENO => #_w1);
   "Shuttle_TCP_Comms_FB_DB_2"(EN := #_w1,   // "Shuttle_TCP_Comms"
                           Enable := "TCP_IP_Shuttle_DB_2".enable,
                           "E-stop" := "L1_OK",
                           TCP_Configuration := "TCP_IP_Shuttle_DB_2".tcpConfig,
                           Shuttle_No := 2,
                           TCP_Diag := "TCP_IP_Shuttle_DB_2".tcpDiagnostics,
                           LCom_Communication_DB := "LCom_Comm_Shuttle_FB_DB_2",
                           Connected => "TCP_IP_Shuttle_DB_2".connected,
                           Busy => "TCP_IP_Shuttle_DB_2".busy,
                           Status => "TCP_IP_Shuttle_DB_2".status,
                           Error => "TCP_IP_Shuttle_DB_2".error,
                           ENO => #_w2);
   IF #_w2 THEN
       "Shuttle_TCP_Comms_FB_DB_3"(Enable := "TCP_IP_Shuttle_DB_3".enable,   // "Shuttle_TCP_Comms"
                               "E-stop" := "L2_OK",
                               TCP_Configuration := "TCP_IP_Shuttle_DB_3".tcpConfig,
                               Shuttle_No := 3,
                               TCP_Diag := "TCP_IP_Shuttle_DB_3".tcpDiagnostics,
                               LCom_Communication_DB := "LCom_Comm_Shuttle_FB_DB_3",
                               Connected => "TCP_IP_Shuttle_DB_3".connected,
                               Busy => "TCP_IP_Shuttle_DB_3".busy,
                               Status => "TCP_IP_Shuttle_DB_3".status,
                               Error => "TCP_IP_Shuttle_DB_3".error);
   END_IF;
   "Shuttle_TCP_Comms_FB_DB_4"(Enable := "TCP_IP_Shuttle_DB_4".enable,   // "Shuttle_TCP_Comms"
                           "E-stop" := "L2_OK",
                           TCP_Configuration := "TCP_IP_Shuttle_DB_4".tcpConfig,
                           Shuttle_No := 4,
                           TCP_Diag := "TCP_IP_Shuttle_DB_4".tcpDiagnostics,
                           LCom_Communication_DB := "LCom_Comm_Shuttle_FB_DB_4",
                           Connected => "TCP_IP_Shuttle_DB_4".connected,
                           Busy => "TCP_IP_Shuttle_DB_4".busy,
                           Status => "TCP_IP_Shuttle_DB_4".status,
                           Error => "TCP_IP_Shuttle_DB_4".error,
                           ENO => #_w3);
   "Shuttle_TCP_Comms_FB_DB_5"(EN := #_w3,   // "Shuttle_TCP_Comms"
                           Enable := "TCP_IP_Shuttle_DB_5".enable,
                           "E-stop" := "L2_OK",
                           TCP_Configuration := "TCP_IP_Shuttle_DB_5".tcpConfig,
                           Shuttle_No := 5,
                           TCP_Diag := "TCP_IP_Shuttle_DB_5".tcpDiagnostics,
                           LCom_Communication_DB := "LCom_Comm_Shuttle_FB_DB_5",
                           Connected => "TCP_IP_Shuttle_DB_5".connected,
                           Busy => "TCP_IP_Shuttle_DB_5".busy,
                           Status => "TCP_IP_Shuttle_DB_5".status,
                           Error => "TCP_IP_Shuttle_DB_5".error,
                           ENO => #_w4);
   IF #_w4 THEN
       "Shuttle_TCP_Comms_FB_DB_6"(Enable := "TCP_IP_Shuttle_DB_6".enable,   // "Shuttle_TCP_Comms"
                               "E-stop" := "L3_OK",
                               TCP_Configuration := "TCP_IP_Shuttle_DB_6".tcpConfig,
                               Shuttle_No := 6,
                               TCP_Diag := "TCP_IP_Shuttle_DB_6".tcpDiagnostics,
                               LCom_Communication_DB := "LCom_Comm_Shuttle_FB_DB_6",
                               Connected => "TCP_IP_Shuttle_DB_6".connected,
                               Busy => "TCP_IP_Shuttle_DB_6".busy,
                               Status => "TCP_IP_Shuttle_DB_6".status,
                               Error => "TCP_IP_Shuttle_DB_6".error);
   END_IF;
   "Shuttle_TCP_Comms_FB_DB_7"(Enable := "TCP_IP_Shuttle_DB_7".enable,   // "Shuttle_TCP_Comms"
                           "E-stop" := "L3_OK",
                           TCP_Configuration := "TCP_IP_Shuttle_DB_7".tcpConfig,
                           Shuttle_No := 7,
                           TCP_Diag := "TCP_IP_Shuttle_DB_7".tcpDiagnostics,
                           LCom_Communication_DB := "LCom_Comm_Shuttle_FB_DB_7",
                           Connected => "TCP_IP_Shuttle_DB_7".connected,
                           Busy => "TCP_IP_Shuttle_DB_7".busy,
                           Status => "TCP_IP_Shuttle_DB_7".status,
                           Error => "TCP_IP_Shuttle_DB_7".error,
                           ENO => #_w5);
   "Shuttle_TCP_Comms_FB_DB_8"(EN := #_w5,   // "Shuttle_TCP_Comms"
                           Enable := "TCP_IP_Shuttle_DB_8".enable,
                           "E-stop" := "L3_OK",
                           TCP_Configuration := "TCP_IP_Shuttle_DB_8".tcpConfig,
                           Shuttle_No := 8,
                           TCP_Diag := "TCP_IP_Shuttle_DB_8".tcpDiagnostics,
                           LCom_Communication_DB := "LCom_Comm_Shuttle_FB_DB_8",
                           Connected => "TCP_IP_Shuttle_DB_8".connected,
                           Busy => "TCP_IP_Shuttle_DB_8".busy,
                           Status => "TCP_IP_Shuttle_DB_8".status,
                           Error => "TCP_IP_Shuttle_DB_8".error,
                           ENO => #_w6);
   IF #_w6 THEN
       "Shuttle_TCP_Comms_FB_DB_9"(Enable := "TCP_IP_Shuttle_DB_9".enable,   // "Shuttle_TCP_Comms"
                               "E-stop" := "L4_OK",
                               TCP_Configuration := "TCP_IP_Shuttle_DB_9".tcpConfig,
                               Shuttle_No := 9,
                               TCP_Diag := "TCP_IP_Shuttle_DB_9".tcpDiagnostics,
                               LCom_Communication_DB := "LCom_Comm_Shuttle_FB_DB_9",
                               Connected => "TCP_IP_Shuttle_DB_9".connected,
                               Busy => "TCP_IP_Shuttle_DB_9".busy,
                               Status => "TCP_IP_Shuttle_DB_9".status,
                               Error => "TCP_IP_Shuttle_DB_9".error);
   END_IF;
   "Shuttle_TCP_Comms_FB_DB_10"(Enable := "TCP_IP_Shuttle_DB_10".enable,   // "Shuttle_TCP_Comms"
                           "E-stop" := "L4_OK",
                           TCP_Configuration := "TCP_IP_Shuttle_DB_10".tcpConfig,
                           Shuttle_No := 10,
                           TCP_Diag := "TCP_IP_Shuttle_DB_10".tcpDiagnostics,
                           LCom_Communication_DB := "LCom_Comm_Shuttle_FB_DB_10",
                           Connected => "TCP_IP_Shuttle_DB_10".connected,
                           Busy => "TCP_IP_Shuttle_DB_10".busy,
                           Status => "TCP_IP_Shuttle_DB_10".status,
                           Error => "TCP_IP_Shuttle_DB_10".error,
                           ENO => #_w7);
   "Shuttle_TCP_Comms_FB_DB_11"(EN := #_w7,   // "Shuttle_TCP_Comms"
                           Enable := "TCP_IP_Shuttle_DB_11".enable,
                           "E-stop" := "L4_OK",
                           TCP_Configuration := "TCP_IP_Shuttle_DB_11".tcpConfig,
                           Shuttle_No := 11,
                           TCP_Diag := "TCP_IP_Shuttle_DB_11".tcpDiagnostics,
                           LCom_Communication_DB := "LCom_Comm_Shuttle_FB_DB_11",
                           Connected => "TCP_IP_Shuttle_DB_11".connected,
                           Busy => "TCP_IP_Shuttle_DB_11".busy,
                           Status => "TCP_IP_Shuttle_DB_11".status,
                           Error => "TCP_IP_Shuttle_DB_11".error,
                           ENO => #_w8);
   IF #_w8 THEN
       "Shuttle_TCP_Comms_FB_DB_12"(Enable := "TCP_IP_Shuttle_DB_12".enable,   // "Shuttle_TCP_Comms"
                               "E-stop" := "L5_OK",
                               TCP_Configuration := "TCP_IP_Shuttle_DB_12".tcpConfig,
                               Shuttle_No := 12,
                               TCP_Diag := "TCP_IP_Shuttle_DB_12".tcpDiagnostics,
                               LCom_Communication_DB := "LCom_Comm_Shuttle_FB_DB_12",
                               Connected => "TCP_IP_Shuttle_DB_12".connected,
                               Busy => "TCP_IP_Shuttle_DB_12".busy,
                               Status => "TCP_IP_Shuttle_DB_12".status,
                               Error => "TCP_IP_Shuttle_DB_12".error);
   END_IF;
   "Shuttle_TCP_Comms_FB_DB_13"(Enable := "TCP_IP_Shuttle_DB_13".enable,   // "Shuttle_TCP_Comms"
                           "E-stop" := "L5_OK",
                           TCP_Configuration := "TCP_IP_Shuttle_DB_13".tcpConfig,
                           Shuttle_No := 13,
                           TCP_Diag := "TCP_IP_Shuttle_DB_13".tcpDiagnostics,
                           LCom_Communication_DB := "LCom_Comm_Shuttle_FB_DB_13",
                           Connected => "TCP_IP_Shuttle_DB_13".connected,
                           Busy => "TCP_IP_Shuttle_DB_13".busy,
                           Status => "TCP_IP_Shuttle_DB_13".status,
                           Error => "TCP_IP_Shuttle_DB_13".error,
                           ENO => #_w9);
   "Shuttle_TCP_Comms_FB_DB_14"(EN := #_w9,   // "Shuttle_TCP_Comms"
                           Enable := "TCP_IP_Shuttle_DB_14".enable,
                           "E-stop" := "L5_OK",
                           TCP_Configuration := "TCP_IP_Shuttle_DB_14".tcpConfig,
                           Shuttle_No := 14,
                           TCP_Diag := "TCP_IP_Shuttle_DB_14".tcpDiagnostics,
                           LCom_Communication_DB := "LCom_Comm_Shuttle_FB_DB_14",
                           Connected => "TCP_IP_Shuttle_DB_14".connected,
                           Busy => "TCP_IP_Shuttle_DB_14".busy,
                           Status => "TCP_IP_Shuttle_DB_14".status,
                           Error => "TCP_IP_Shuttle_DB_14".error,
                           ENO => #_w10);
   IF #_w10 THEN
       "Shuttle_TCP_Comms_FB_DB_15"(Enable := "TCP_IP_Shuttle_DB_15".enable,   // "Shuttle_TCP_Comms"
                               "E-stop" := "L6_OK",
                               TCP_Configuration := "TCP_IP_Shuttle_DB_15".tcpConfig,
                               Shuttle_No := 15,
                               TCP_Diag := "TCP_IP_Shuttle_DB_15".tcpDiagnostics,
                               LCom_Communication_DB := "LCom_Comm_Shuttle_FB_DB_15",
                               Connected => "TCP_IP_Shuttle_DB_15".connected,
                               Busy => "TCP_IP_Shuttle_DB_15".busy,
                               Status => "TCP_IP_Shuttle_DB_15".status,
                               Error => "TCP_IP_Shuttle_DB_15".error);
   END_IF;
   "Shuttle_TCP_Comms_FB_DB_16"(Enable := "TCP_IP_Shuttle_DB_16".enable,   // "Shuttle_TCP_Comms"
                           "E-stop" := "L6_OK",
                           TCP_Configuration := "TCP_IP_Shuttle_DB_16".tcpConfig,
                           Shuttle_No := 16,
                           TCP_Diag := "TCP_IP_Shuttle_DB_16".tcpDiagnostics,
                           LCom_Communication_DB := "LCom_Comm_Shuttle_FB_DB_16",
                           Connected => "TCP_IP_Shuttle_DB_16".connected,
                           Busy => "TCP_IP_Shuttle_DB_16".busy,
                           Status => "TCP_IP_Shuttle_DB_16".status,
                           Error => "TCP_IP_Shuttle_DB_16".error,
                           ENO => #_w11);
   "Shuttle_TCP_Comms_FB_DB_17"(EN := #_w11,   // "Shuttle_TCP_Comms"
                           Enable := "TCP_IP_Shuttle_DB_17".enable,
                           "E-stop" := "L6_OK",
                           TCP_Configuration := "TCP_IP_Shuttle_DB_17".tcpConfig,
                           Shuttle_No := 17,
                           TCP_Diag := "TCP_IP_Shuttle_DB_17".tcpDiagnostics,
                           LCom_Communication_DB := "LCom_Comm_Shuttle_FB_DB_17",
                           Connected => "TCP_IP_Shuttle_DB_17".connected,
                           Busy => "TCP_IP_Shuttle_DB_17".busy,
                           Status => "TCP_IP_Shuttle_DB_17".status,
                           Error => "TCP_IP_Shuttle_DB_17".error,
                           ENO => #_w12);
   IF #_w12 THEN
       "Shuttle_TCP_Comms_FB_DB_18"(Enable := "TCP_IP_Shuttle_DB_18".enable,   // "Shuttle_TCP_Comms"
                               "E-stop" := "L7_OK",
                               TCP_Configuration := "TCP_IP_Shuttle_DB_18".tcpConfig,
                               Shuttle_No := 18,
                               TCP_Diag := "TCP_IP_Shuttle_DB_18".tcpDiagnostics,
                               LCom_Communication_DB := "LCom_Comm_Shuttle_FB_DB_18",
                               Connected => "TCP_IP_Shuttle_DB_18".connected,
                               Busy => "TCP_IP_Shuttle_DB_18".busy,
                               Status => "TCP_IP_Shuttle_DB_18".status,
                               Error => "TCP_IP_Shuttle_DB_18".error);
   END_IF;
   "Shuttle_TCP_Comms_FB_DB_19"(Enable := "TCP_IP_Shuttle_DB_19".enable,   // "Shuttle_TCP_Comms"
                           "E-stop" := "L7_OK",
                           TCP_Configuration := "TCP_IP_Shuttle_DB_19".tcpConfig,
                           Shuttle_No := 19,
                           TCP_Diag := "TCP_IP_Shuttle_DB_19".tcpDiagnostics,
                           LCom_Communication_DB := "LCom_Comm_Shuttle_FB_DB_19",
                           Connected => "TCP_IP_Shuttle_DB_19".connected,
                           Busy => "TCP_IP_Shuttle_DB_19".busy,
                           Status => "TCP_IP_Shuttle_DB_19".status,
                           Error => "TCP_IP_Shuttle_DB_19".error,
                           ENO => #_w13);
   "Shuttle_TCP_Comms_FB_DB_20"(EN := #_w13,   // "Shuttle_TCP_Comms"
                           Enable := "TCP_IP_Shuttle_DB_20".enable,
                           "E-stop" := "L7_OK",
                           TCP_Configuration := "TCP_IP_Shuttle_DB_20".tcpConfig,
                           Shuttle_No := 20,
                           TCP_Diag := "TCP_IP_Shuttle_DB_20".tcpDiagnostics,
                           LCom_Communication_DB := "LCom_Comm_Shuttle_FB_DB_20",
                           Connected => "TCP_IP_Shuttle_DB_20".connected,
                           Busy => "TCP_IP_Shuttle_DB_20".busy,
                           Status => "TCP_IP_Shuttle_DB_20".status,
                           Error => "TCP_IP_Shuttle_DB_20".error,
                           ENO => #_w14);
   IF #_w14 THEN
       "Shuttle_TCP_Comms_FB_DB_21"(Enable := "TCP_IP_Shuttle_DB_21".enable,   // "Shuttle_TCP_Comms"
                               "E-stop" := "L8_OK",
                               TCP_Configuration := "TCP_IP_Shuttle_DB_21".tcpConfig,
                               Shuttle_No := 21,
                               TCP_Diag := "TCP_IP_Shuttle_DB_21".tcpDiagnostics,
                               LCom_Communication_DB := "LCom_Comm_Shuttle_FB_DB_21",
                               Connected => "TCP_IP_Shuttle_DB_21".connected,
                               Busy => "TCP_IP_Shuttle_DB_21".busy,
                               Status => "TCP_IP_Shuttle_DB_21".status,
                               Error => "TCP_IP_Shuttle_DB_21".error);
   END_IF;
   "Shuttle_TCP_Comms_FB_DB_22"(Enable := "TCP_IP_Shuttle_DB_22".enable,   // "Shuttle_TCP_Comms"
                           "E-stop" := "L8_OK",
                           TCP_Configuration := "TCP_IP_Shuttle_DB_22".tcpConfig,
                           Shuttle_No := 22,
                           TCP_Diag := "TCP_IP_Shuttle_DB_22".tcpDiagnostics,
                           LCom_Communication_DB := "LCom_Comm_Shuttle_FB_DB_22",
                           Connected => "TCP_IP_Shuttle_DB_22".connected,
                           Busy => "TCP_IP_Shuttle_DB_22".busy,
                           Status => "TCP_IP_Shuttle_DB_22".status,
                           Error => "TCP_IP_Shuttle_DB_22".error,
                           ENO => #_w15);
   IF #_w15 THEN
       "Shuttle_TCP_Comms_FB_DB_23"(Enable := "TCP_IP_Shuttle_DB_23".enable,   // "Shuttle_TCP_Comms"
                               "E-stop" := "L8_OK",
                               TCP_Configuration := "TCP_IP_Shuttle_DB_23".tcpConfig,
                               Shuttle_No := 23,
                               TCP_Diag := "TCP_IP_Shuttle_DB_23".tcpDiagnostics,
                               LCom_Communication_DB := "LCom_Comm_Shuttle_FB_DB_23",
                               Connected => "TCP_IP_Shuttle_DB_23".connected,
                               Busy => "TCP_IP_Shuttle_DB_23".busy,
                               Status => "TCP_IP_Shuttle_DB_23".status,
                               Error => "TCP_IP_Shuttle_DB_23".error);
   END_IF;
END_REGION

REGION Network 50: GATE STATIONS SYSTEMS 1,2 (Gates 1 and 2)
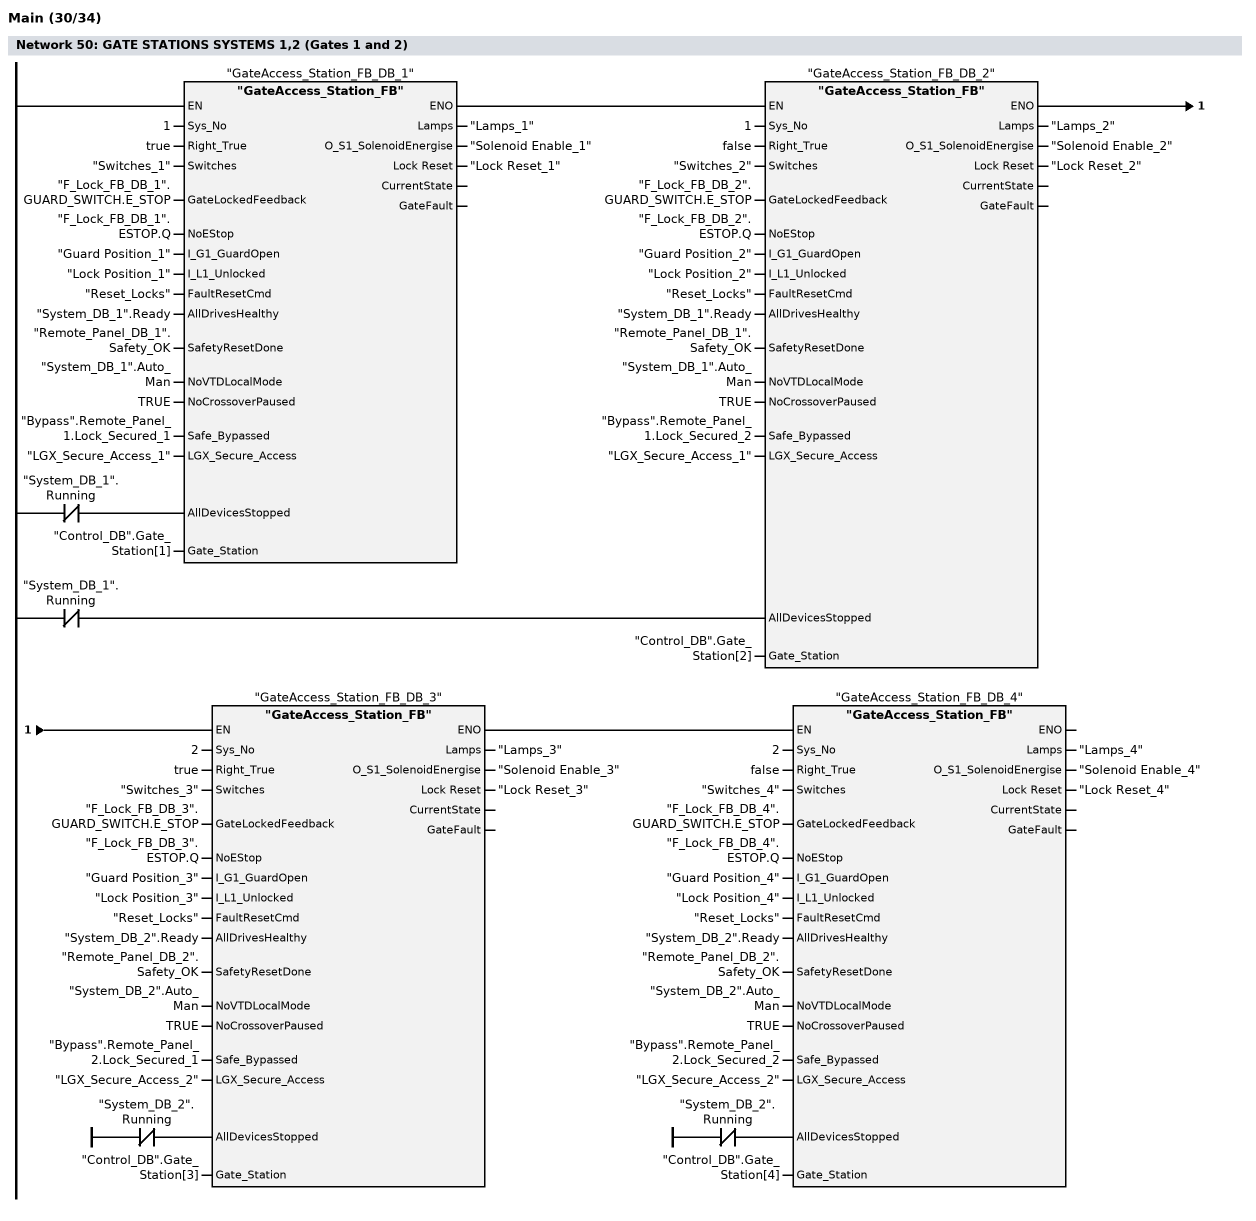
   RUNG wire#powerrail
      "GateAccess_Station_FB_DB_1"(AllDevicesStopped := wire#w1, Sys_No := 1, Right_True := true, Switches := "Switches_1", GateLockedFeedback := "F_Lock_FB_DB_1".GUARD_SWITCH.E_STOP, NoEStop := "F_Lock_FB_DB_1".ESTOP.Q, I_G1_GuardOpen := "Guard Position_1", I_L1_Unlocked := "Lock Position_1", FaultResetCmd := "Reset_Locks", AllDrivesHealthy := "System_DB_1".Ready, SafetyResetDone := "Remote_Panel_DB_1".Safety_OK, NoVTDLocalMode := "System_DB_1".Auto_Man, NoCrossoverPaused := TRUE, Safe_Bypassed := "Bypass".Remote_Panel_1.Lock_Secured_1, LGX_Secure_Access := "LGX_Secure_Access_1", Gate_Station := "Control_DB".Gate_Station[1], Lamps => "Lamps_1", O_S1_SolenoidEnergise => "Solenoid Enable_1", "Lock Reset" => "Lock Reset_1", CurrentState =>, GateFault =>)
      "GateAccess_Station_FB_DB_2"(AllDevicesStopped := wire#w2, Sys_No := 1, Right_True := false, Switches := "Switches_2", GateLockedFeedback := "F_Lock_FB_DB_2".GUARD_SWITCH.E_STOP, NoEStop := "F_Lock_FB_DB_2".ESTOP.Q, I_G1_GuardOpen := "Guard Position_2", I_L1_Unlocked := "Lock Position_2", FaultResetCmd := "Reset_Locks", AllDrivesHealthy := "System_DB_1".Ready, SafetyResetDone := "Remote_Panel_DB_1".Safety_OK, NoVTDLocalMode := "System_DB_1".Auto_Man, NoCrossoverPaused := TRUE, Safe_Bypassed := "Bypass".Remote_Panel_1.Lock_Secured_2, LGX_Secure_Access := "LGX_Secure_Access_1", Gate_Station := "Control_DB".Gate_Station[2], Lamps => "Lamps_2", O_S1_SolenoidEnergise => "Solenoid Enable_2", "Lock Reset" => "Lock Reset_2", CurrentState =>, GateFault =>)
      "GateAccess_Station_FB_DB_3"(AllDevicesStopped := wire#w3, Sys_No := 2, Right_True := true, Switches := "Switches_3", GateLockedFeedback := "F_Lock_FB_DB_3".GUARD_SWITCH.E_STOP, NoEStop := "F_Lock_FB_DB_3".ESTOP.Q, I_G1_GuardOpen := "Guard Position_3", I_L1_Unlocked := "Lock Position_3", FaultResetCmd := "Reset_Locks", AllDrivesHealthy := "System_DB_2".Ready, SafetyResetDone := "Remote_Panel_DB_2".Safety_OK, NoVTDLocalMode := "System_DB_2".Auto_Man, NoCrossoverPaused := TRUE, Safe_Bypassed := "Bypass".Remote_Panel_2.Lock_Secured_1, LGX_Secure_Access := "LGX_Secure_Access_2", Gate_Station := "Control_DB".Gate_Station[3], Lamps => "Lamps_3", O_S1_SolenoidEnergise => "Solenoid Enable_3", "Lock Reset" => "Lock Reset_3", CurrentState =>, GateFault =>)
      "GateAccess_Station_FB_DB_4"(AllDevicesStopped := wire#w4, Sys_No := 2, Right_True := false, Switches := "Switches_4", GateLockedFeedback := "F_Lock_FB_DB_4".GUARD_SWITCH.E_STOP, NoEStop := "F_Lock_FB_DB_4".ESTOP.Q, I_G1_GuardOpen := "Guard Position_4", I_L1_Unlocked := "Lock Position_4", FaultResetCmd := "Reset_Locks", AllDrivesHealthy := "System_DB_2".Ready, SafetyResetDone := "Remote_Panel_DB_2".Safety_OK, NoVTDLocalMode := "System_DB_2".Auto_Man, NoCrossoverPaused := TRUE, Safe_Bypassed := "Bypass".Remote_Panel_2.Lock_Secured_2, LGX_Secure_Access := "LGX_Secure_Access_2", Gate_Station := "Control_DB".Gate_Station[4], Lamps => "Lamps_4", O_S1_SolenoidEnergise => "Solenoid Enable_4", "Lock Reset" => "Lock Reset_4", CurrentState =>, GateFault =>)
   END_RUNG
   RUNG wire#powerrail
      I_Contact( "System_DB_1".Running )
   END_RUNG wire#w1
   RUNG wire#powerrail
      I_Contact( "System_DB_1".Running )
   END_RUNG wire#w2
   RUNG wire#powerrail
      I_Contact( "System_DB_2".Running )
   END_RUNG wire#w3
   RUNG wire#powerrail
      I_Contact( "System_DB_2".Running )
   END_RUNG wire#w4
   // the same network as SCL:
   "GateAccess_Station_FB_DB_1"(Sys_No := 1,   // "GateAccess_Station_FB"
                           Right_True := true,
                           Switches := "Switches_1",
                           GateLockedFeedback := "F_Lock_FB_DB_1".GUARD_SWITCH.E_STOP,
                           NoEStop := "F_Lock_FB_DB_1".ESTOP.Q,
                           I_G1_GuardOpen := "Guard Position_1",
                           I_L1_Unlocked := "Lock Position_1",
                           FaultResetCmd := "Reset_Locks",
                           AllDrivesHealthy := "System_DB_1".Ready,
                           SafetyResetDone := "Remote_Panel_DB_1".Safety_OK,
                           NoVTDLocalMode := "System_DB_1".Auto_Man,
                           NoCrossoverPaused := TRUE,
                           Safe_Bypassed := "Bypass".Remote_Panel_1.Lock_Secured_1,
                           LGX_Secure_Access := "LGX_Secure_Access_1",
                           AllDevicesStopped := NOT "System_DB_1".Running,
                           Gate_Station := "Control_DB".Gate_Station[1],
                           Lamps => "Lamps_1",
                           O_S1_SolenoidEnergise => "Solenoid Enable_1",
                           "Lock Reset" => "Lock Reset_1",
                           ENO => #_w1);
   "GateAccess_Station_FB_DB_2"(EN := #_w1,   // "GateAccess_Station_FB"
                           Sys_No := 1,
                           Right_True := false,
                           Switches := "Switches_2",
                           GateLockedFeedback := "F_Lock_FB_DB_2".GUARD_SWITCH.E_STOP,
                           NoEStop := "F_Lock_FB_DB_2".ESTOP.Q,
                           I_G1_GuardOpen := "Guard Position_2",
                           I_L1_Unlocked := "Lock Position_2",
                           FaultResetCmd := "Reset_Locks",
                           AllDrivesHealthy := "System_DB_1".Ready,
                           SafetyResetDone := "Remote_Panel_DB_1".Safety_OK,
                           NoVTDLocalMode := "System_DB_1".Auto_Man,
                           NoCrossoverPaused := TRUE,
                           Safe_Bypassed := "Bypass".Remote_Panel_1.Lock_Secured_2,
                           LGX_Secure_Access := "LGX_Secure_Access_1",
                           AllDevicesStopped := NOT "System_DB_1".Running,
                           Gate_Station := "Control_DB".Gate_Station[2],
                           Lamps => "Lamps_2",
                           O_S1_SolenoidEnergise => "Solenoid Enable_2",
                           "Lock Reset" => "Lock Reset_2",
                           ENO => #_w2);
   "GateAccess_Station_FB_DB_3"(EN := #_w2,   // "GateAccess_Station_FB"
                           Sys_No := 2,
                           Right_True := true,
                           Switches := "Switches_3",
                           GateLockedFeedback := "F_Lock_FB_DB_3".GUARD_SWITCH.E_STOP,
                           NoEStop := "F_Lock_FB_DB_3".ESTOP.Q,
                           I_G1_GuardOpen := "Guard Position_3",
                           I_L1_Unlocked := "Lock Position_3",
                           FaultResetCmd := "Reset_Locks",
                           AllDrivesHealthy := "System_DB_2".Ready,
                           SafetyResetDone := "Remote_Panel_DB_2".Safety_OK,
                           NoVTDLocalMode := "System_DB_2".Auto_Man,
                           NoCrossoverPaused := TRUE,
                           Safe_Bypassed := "Bypass".Remote_Panel_2.Lock_Secured_1,
                           LGX_Secure_Access := "LGX_Secure_Access_2",
                           AllDevicesStopped := NOT "System_DB_2".Running,
                           Gate_Station := "Control_DB".Gate_Station[3],
                           Lamps => "Lamps_3",
                           O_S1_SolenoidEnergise => "Solenoid Enable_3",
                           "Lock Reset" => "Lock Reset_3",
                           ENO => #_w3);
   IF #_w3 THEN
       "GateAccess_Station_FB_DB_4"(Sys_No := 2,   // "GateAccess_Station_FB"
                               Right_True := false,
                               Switches := "Switches_4",
                               GateLockedFeedback := "F_Lock_FB_DB_4".GUARD_SWITCH.E_STOP,
                               NoEStop := "F_Lock_FB_DB_4".ESTOP.Q,
                               I_G1_GuardOpen := "Guard Position_4",
                               I_L1_Unlocked := "Lock Position_4",
                               FaultResetCmd := "Reset_Locks",
                               AllDrivesHealthy := "System_DB_2".Ready,
                               SafetyResetDone := "Remote_Panel_DB_2".Safety_OK,
                               NoVTDLocalMode := "System_DB_2".Auto_Man,
                               NoCrossoverPaused := TRUE,
                               Safe_Bypassed := "Bypass".Remote_Panel_2.Lock_Secured_2,
                               LGX_Secure_Access := "LGX_Secure_Access_2",
                               AllDevicesStopped := NOT "System_DB_2".Running,
                               Gate_Station := "Control_DB".Gate_Station[4],
                               Lamps => "Lamps_4",
                               O_S1_SolenoidEnergise => "Solenoid Enable_4",
                               "Lock Reset" => "Lock Reset_4");
   END_IF;
END_REGION

REGION Network 51: GATE STATIONS SYSTEMS 3 (Gates 1 and 2)
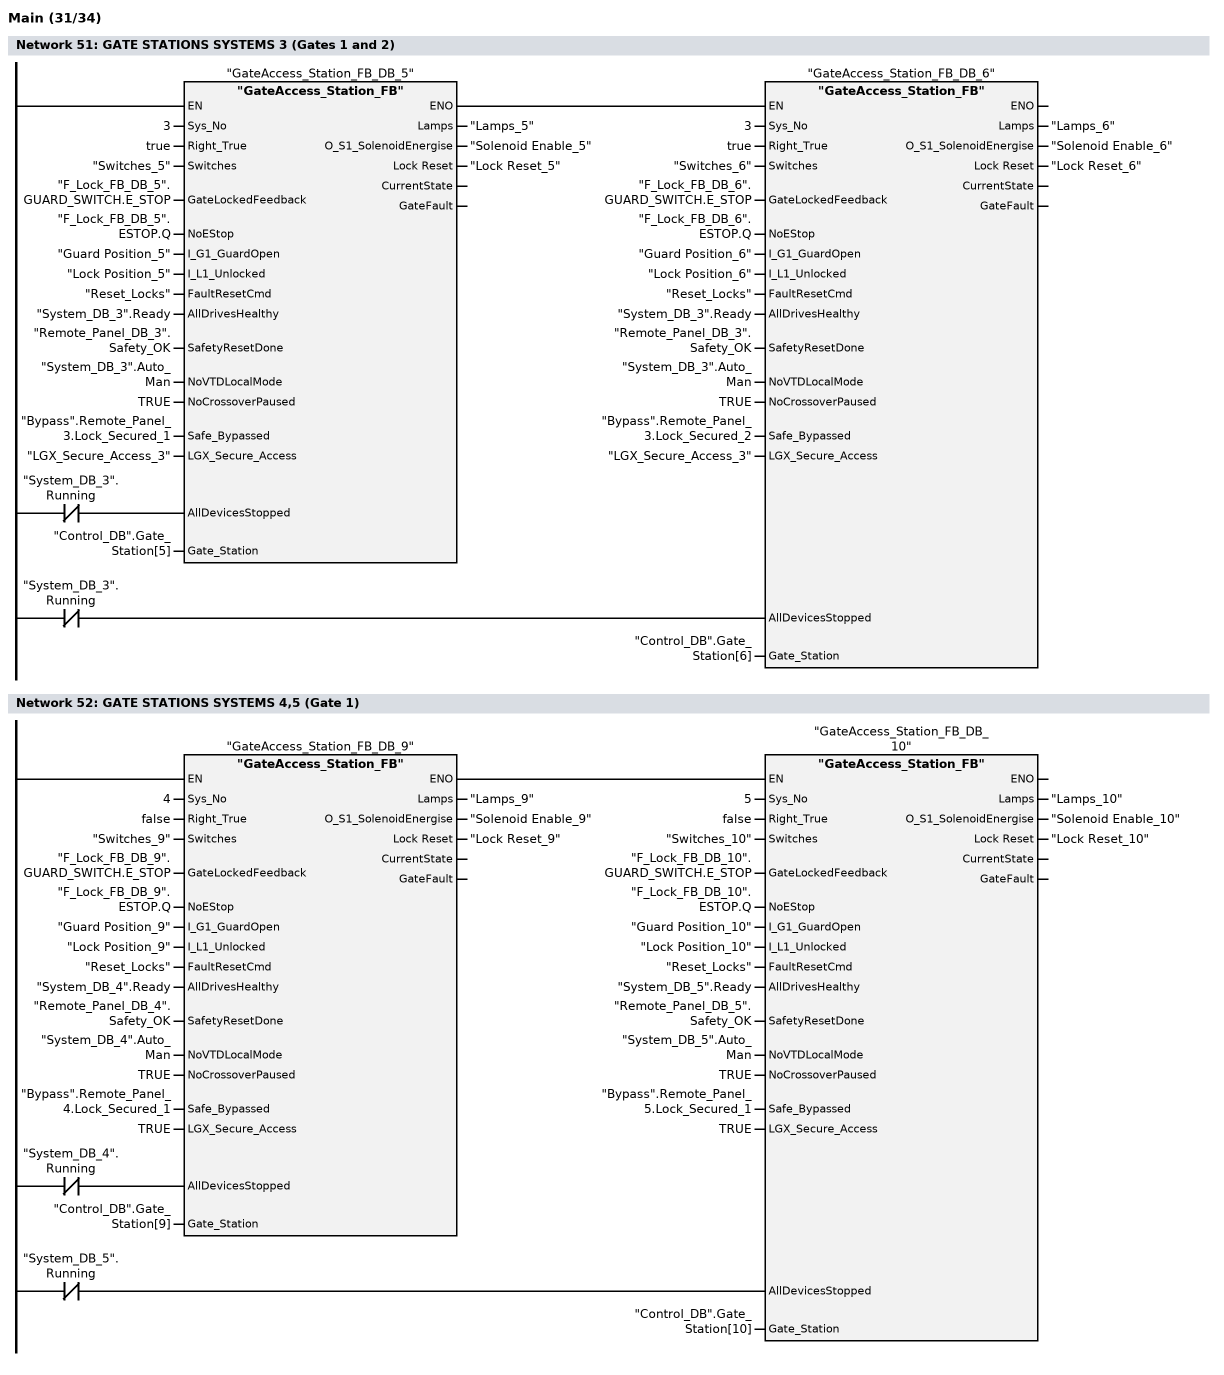
   RUNG wire#powerrail
      "GateAccess_Station_FB_DB_5"(AllDevicesStopped := wire#w1, Sys_No := 3, Right_True := true, Switches := "Switches_5", GateLockedFeedback := "F_Lock_FB_DB_5".GUARD_SWITCH.E_STOP, NoEStop := "F_Lock_FB_DB_5".ESTOP.Q, I_G1_GuardOpen := "Guard Position_5", I_L1_Unlocked := "Lock Position_5", FaultResetCmd := "Reset_Locks", AllDrivesHealthy := "System_DB_3".Ready, SafetyResetDone := "Remote_Panel_DB_3".Safety_OK, NoVTDLocalMode := "System_DB_3".Auto_Man, NoCrossoverPaused := TRUE, Safe_Bypassed := "Bypass".Remote_Panel_3.Lock_Secured_1, LGX_Secure_Access := "LGX_Secure_Access_3", Gate_Station := "Control_DB".Gate_Station[5], Lamps => "Lamps_5", O_S1_SolenoidEnergise => "Solenoid Enable_5", "Lock Reset" => "Lock Reset_5", CurrentState =>, GateFault =>)
      "GateAccess_Station_FB_DB_6"(AllDevicesStopped := wire#w2, Sys_No := 3, Right_True := true, Switches := "Switches_6", GateLockedFeedback := "F_Lock_FB_DB_6".GUARD_SWITCH.E_STOP, NoEStop := "F_Lock_FB_DB_6".ESTOP.Q, I_G1_GuardOpen := "Guard Position_6", I_L1_Unlocked := "Lock Position_6", FaultResetCmd := "Reset_Locks", AllDrivesHealthy := "System_DB_3".Ready, SafetyResetDone := "Remote_Panel_DB_3".Safety_OK, NoVTDLocalMode := "System_DB_3".Auto_Man, NoCrossoverPaused := TRUE, Safe_Bypassed := "Bypass".Remote_Panel_3.Lock_Secured_2, LGX_Secure_Access := "LGX_Secure_Access_3", Gate_Station := "Control_DB".Gate_Station[6], Lamps => "Lamps_6", O_S1_SolenoidEnergise => "Solenoid Enable_6", "Lock Reset" => "Lock Reset_6", CurrentState =>, GateFault =>)
   END_RUNG
   RUNG wire#powerrail
      I_Contact( "System_DB_3".Running )
   END_RUNG wire#w1
   RUNG wire#powerrail
      I_Contact( "System_DB_3".Running )
   END_RUNG wire#w2
   // the same network as SCL:
   "GateAccess_Station_FB_DB_5"(Sys_No := 3,   // "GateAccess_Station_FB"
                           Right_True := true,
                           Switches := "Switches_5",
                           GateLockedFeedback := "F_Lock_FB_DB_5".GUARD_SWITCH.E_STOP,
                           NoEStop := "F_Lock_FB_DB_5".ESTOP.Q,
                           I_G1_GuardOpen := "Guard Position_5",
                           I_L1_Unlocked := "Lock Position_5",
                           FaultResetCmd := "Reset_Locks",
                           AllDrivesHealthy := "System_DB_3".Ready,
                           SafetyResetDone := "Remote_Panel_DB_3".Safety_OK,
                           NoVTDLocalMode := "System_DB_3".Auto_Man,
                           NoCrossoverPaused := TRUE,
                           Safe_Bypassed := "Bypass".Remote_Panel_3.Lock_Secured_1,
                           LGX_Secure_Access := "LGX_Secure_Access_3",
                           AllDevicesStopped := NOT "System_DB_3".Running,
                           Gate_Station := "Control_DB".Gate_Station[5],
                           Lamps => "Lamps_5",
                           O_S1_SolenoidEnergise => "Solenoid Enable_5",
                           "Lock Reset" => "Lock Reset_5",
                           ENO => #_w1);
   IF #_w1 THEN
       "GateAccess_Station_FB_DB_6"(Sys_No := 3,   // "GateAccess_Station_FB"
                               Right_True := true,
                               Switches := "Switches_6",
                               GateLockedFeedback := "F_Lock_FB_DB_6".GUARD_SWITCH.E_STOP,
                               NoEStop := "F_Lock_FB_DB_6".ESTOP.Q,
                               I_G1_GuardOpen := "Guard Position_6",
                               I_L1_Unlocked := "Lock Position_6",
                               FaultResetCmd := "Reset_Locks",
                               AllDrivesHealthy := "System_DB_3".Ready,
                               SafetyResetDone := "Remote_Panel_DB_3".Safety_OK,
                               NoVTDLocalMode := "System_DB_3".Auto_Man,
                               NoCrossoverPaused := TRUE,
                               Safe_Bypassed := "Bypass".Remote_Panel_3.Lock_Secured_2,
                               LGX_Secure_Access := "LGX_Secure_Access_3",
                               AllDevicesStopped := NOT "System_DB_3".Running,
                               Gate_Station := "Control_DB".Gate_Station[6],
                               Lamps => "Lamps_6",
                               O_S1_SolenoidEnergise => "Solenoid Enable_6",
                               "Lock Reset" => "Lock Reset_6");
   END_IF;
END_REGION

REGION Network 52: GATE STATIONS SYSTEMS 4,5 (Gate 1)
   RUNG wire#powerrail
      "GateAccess_Station_FB_DB_9"(AllDevicesStopped := wire#w1, Sys_No := 4, Right_True := false, Switches := "Switches_9", GateLockedFeedback := "F_Lock_FB_DB_9".GUARD_SWITCH.E_STOP, NoEStop := "F_Lock_FB_DB_9".ESTOP.Q, I_G1_GuardOpen := "Guard Position_9", I_L1_Unlocked := "Lock Position_9", FaultResetCmd := "Reset_Locks", AllDrivesHealthy := "System_DB_4".Ready, SafetyResetDone := "Remote_Panel_DB_4".Safety_OK, NoVTDLocalMode := "System_DB_4".Auto_Man, NoCrossoverPaused := TRUE, Safe_Bypassed := "Bypass".Remote_Panel_4.Lock_Secured_1, LGX_Secure_Access := TRUE, Gate_Station := "Control_DB".Gate_Station[9], Lamps => "Lamps_9", O_S1_SolenoidEnergise => "Solenoid Enable_9", "Lock Reset" => "Lock Reset_9", CurrentState =>, GateFault =>)
      "GateAccess_Station_FB_DB_10"(AllDevicesStopped := wire#w2, Sys_No := 5, Right_True := false, Switches := "Switches_10", GateLockedFeedback := "F_Lock_FB_DB_10".GUARD_SWITCH.E_STOP, NoEStop := "F_Lock_FB_DB_10".ESTOP.Q, I_G1_GuardOpen := "Guard Position_10", I_L1_Unlocked := "Lock Position_10", FaultResetCmd := "Reset_Locks", AllDrivesHealthy := "System_DB_5".Ready, SafetyResetDone := "Remote_Panel_DB_5".Safety_OK, NoVTDLocalMode := "System_DB_5".Auto_Man, NoCrossoverPaused := TRUE, Safe_Bypassed := "Bypass".Remote_Panel_5.Lock_Secured_1, LGX_Secure_Access := TRUE, Gate_Station := "Control_DB".Gate_Station[10], Lamps => "Lamps_10", O_S1_SolenoidEnergise => "Solenoid Enable_10", "Lock Reset" => "Lock Reset_10", CurrentState =>, GateFault =>)
   END_RUNG
   RUNG wire#powerrail
      I_Contact( "System_DB_4".Running )
   END_RUNG wire#w1
   RUNG wire#powerrail
      I_Contact( "System_DB_5".Running )
   END_RUNG wire#w2
   // the same network as SCL:
   "GateAccess_Station_FB_DB_9"(Sys_No := 4,   // "GateAccess_Station_FB"
                           Right_True := false,
                           Switches := "Switches_9",
                           GateLockedFeedback := "F_Lock_FB_DB_9".GUARD_SWITCH.E_STOP,
                           NoEStop := "F_Lock_FB_DB_9".ESTOP.Q,
                           I_G1_GuardOpen := "Guard Position_9",
                           I_L1_Unlocked := "Lock Position_9",
                           FaultResetCmd := "Reset_Locks",
                           AllDrivesHealthy := "System_DB_4".Ready,
                           SafetyResetDone := "Remote_Panel_DB_4".Safety_OK,
                           NoVTDLocalMode := "System_DB_4".Auto_Man,
                           NoCrossoverPaused := TRUE,
                           Safe_Bypassed := "Bypass".Remote_Panel_4.Lock_Secured_1,
                           LGX_Secure_Access := TRUE,
                           AllDevicesStopped := NOT "System_DB_4".Running,
                           Gate_Station := "Control_DB".Gate_Station[9],
                           Lamps => "Lamps_9",
                           O_S1_SolenoidEnergise => "Solenoid Enable_9",
                           "Lock Reset" => "Lock Reset_9",
                           ENO => #_w1);
   IF #_w1 THEN
       "GateAccess_Station_FB_DB_10"(Sys_No := 5,   // "GateAccess_Station_FB"
                               Right_True := false,
                               Switches := "Switches_10",
                               GateLockedFeedback := "F_Lock_FB_DB_10".GUARD_SWITCH.E_STOP,
                               NoEStop := "F_Lock_FB_DB_10".ESTOP.Q,
                               I_G1_GuardOpen := "Guard Position_10",
                               I_L1_Unlocked := "Lock Position_10",
                               FaultResetCmd := "Reset_Locks",
                               AllDrivesHealthy := "System_DB_5".Ready,
                               SafetyResetDone := "Remote_Panel_DB_5".Safety_OK,
                               NoVTDLocalMode := "System_DB_5".Auto_Man,
                               NoCrossoverPaused := TRUE,
                               Safe_Bypassed := "Bypass".Remote_Panel_5.Lock_Secured_1,
                               LGX_Secure_Access := TRUE,
                               AllDevicesStopped := NOT "System_DB_5".Running,
                               Gate_Station := "Control_DB".Gate_Station[10],
                               Lamps => "Lamps_10",
                               O_S1_SolenoidEnergise => "Solenoid Enable_10",
                               "Lock Reset" => "Lock Reset_10");
   END_IF;
END_REGION

REGION Network 53: Gate Stations Left and Right, Level 1 and Level 2
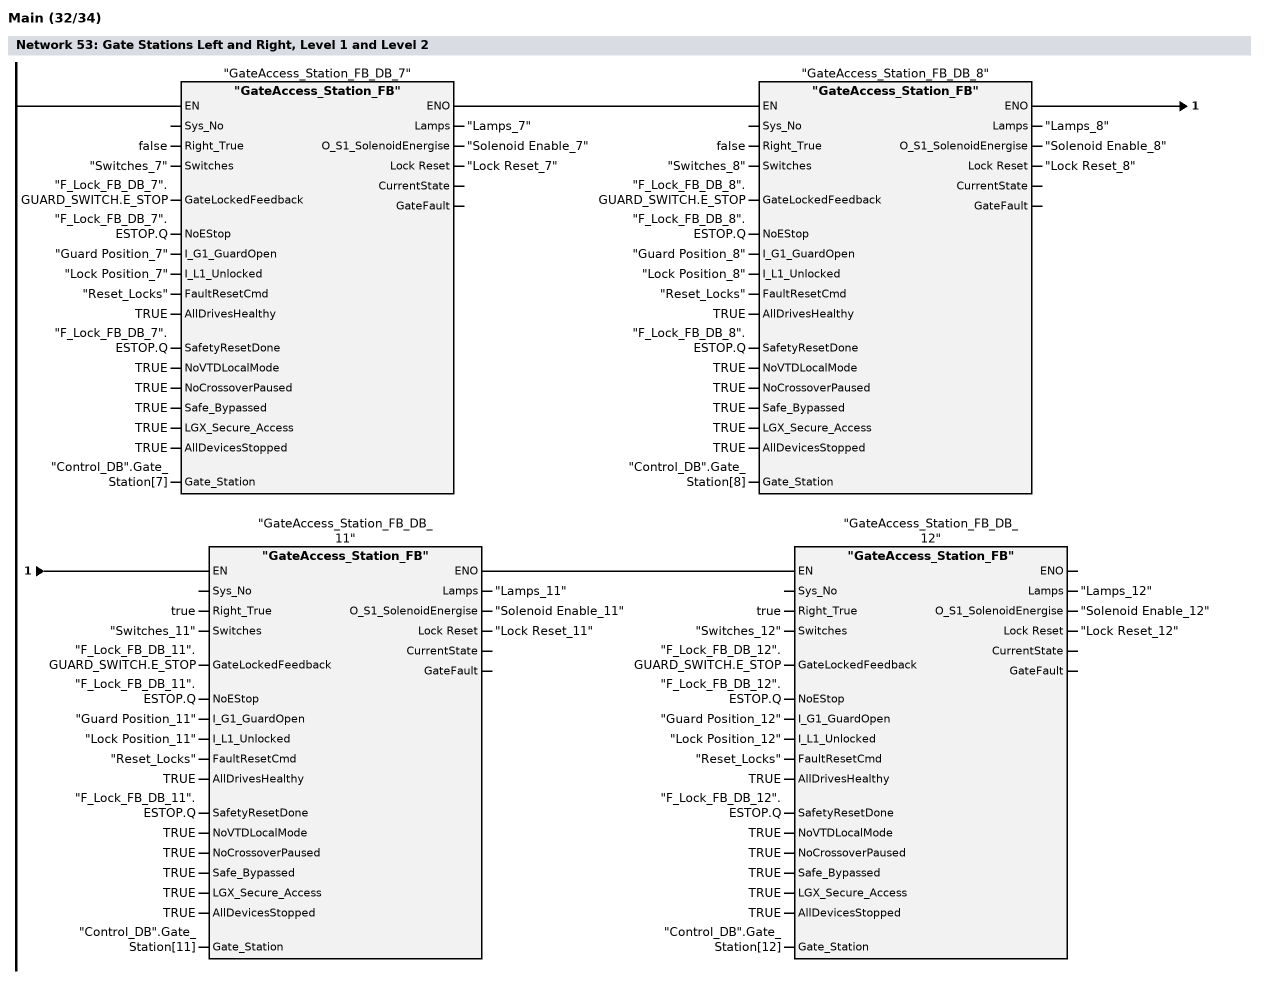
   RUNG wire#powerrail
      "GateAccess_Station_FB_DB_7"(Sys_No :=, Right_True := false, Switches := "Switches_7", GateLockedFeedback := "F_Lock_FB_DB_7".GUARD_SWITCH.E_STOP, NoEStop := "F_Lock_FB_DB_7".ESTOP.Q, I_G1_GuardOpen := "Guard Position_7", I_L1_Unlocked := "Lock Position_7", FaultResetCmd := "Reset_Locks", AllDrivesHealthy := TRUE, SafetyResetDone := "F_Lock_FB_DB_7".ESTOP.Q, NoVTDLocalMode := TRUE, NoCrossoverPaused := TRUE, Safe_Bypassed := TRUE, LGX_Secure_Access := TRUE, AllDevicesStopped := TRUE, Gate_Station := "Control_DB".Gate_Station[7], Lamps => "Lamps_7", O_S1_SolenoidEnergise => "Solenoid Enable_7", "Lock Reset" => "Lock Reset_7", CurrentState =>, GateFault =>)
      "GateAccess_Station_FB_DB_8"(Sys_No :=, Right_True := false, Switches := "Switches_8", GateLockedFeedback := "F_Lock_FB_DB_8".GUARD_SWITCH.E_STOP, NoEStop := "F_Lock_FB_DB_8".ESTOP.Q, I_G1_GuardOpen := "Guard Position_8", I_L1_Unlocked := "Lock Position_8", FaultResetCmd := "Reset_Locks", AllDrivesHealthy := TRUE, SafetyResetDone := "F_Lock_FB_DB_8".ESTOP.Q, NoVTDLocalMode := TRUE, NoCrossoverPaused := TRUE, Safe_Bypassed := TRUE, LGX_Secure_Access := TRUE, AllDevicesStopped := TRUE, Gate_Station := "Control_DB".Gate_Station[8], Lamps => "Lamps_8", O_S1_SolenoidEnergise => "Solenoid Enable_8", "Lock Reset" => "Lock Reset_8", CurrentState =>, GateFault =>)
      "GateAccess_Station_FB_DB_11"(Sys_No :=, Right_True := true, Switches := "Switches_11", GateLockedFeedback := "F_Lock_FB_DB_11".GUARD_SWITCH.E_STOP, NoEStop := "F_Lock_FB_DB_11".ESTOP.Q, I_G1_GuardOpen := "Guard Position_11", I_L1_Unlocked := "Lock Position_11", FaultResetCmd := "Reset_Locks", AllDrivesHealthy := TRUE, SafetyResetDone := "F_Lock_FB_DB_11".ESTOP.Q, NoVTDLocalMode := TRUE, NoCrossoverPaused := TRUE, Safe_Bypassed := TRUE, LGX_Secure_Access := TRUE, AllDevicesStopped := TRUE, Gate_Station := "Control_DB".Gate_Station[11], Lamps => "Lamps_11", O_S1_SolenoidEnergise => "Solenoid Enable_11", "Lock Reset" => "Lock Reset_11", CurrentState =>, GateFault =>)
      "GateAccess_Station_FB_DB_12"(Sys_No :=, Right_True := true, Switches := "Switches_12", GateLockedFeedback := "F_Lock_FB_DB_12".GUARD_SWITCH.E_STOP, NoEStop := "F_Lock_FB_DB_12".ESTOP.Q, I_G1_GuardOpen := "Guard Position_12", I_L1_Unlocked := "Lock Position_12", FaultResetCmd := "Reset_Locks", AllDrivesHealthy := TRUE, SafetyResetDone := "F_Lock_FB_DB_12".ESTOP.Q, NoVTDLocalMode := TRUE, NoCrossoverPaused := TRUE, Safe_Bypassed := TRUE, LGX_Secure_Access := TRUE, AllDevicesStopped := TRUE, Gate_Station := "Control_DB".Gate_Station[12], Lamps => "Lamps_12", O_S1_SolenoidEnergise => "Solenoid Enable_12", "Lock Reset" => "Lock Reset_12", CurrentState =>, GateFault =>)
   END_RUNG
   // the same network as SCL:
   "GateAccess_Station_FB_DB_7"(Right_True := false,   // "GateAccess_Station_FB"
                           Switches := "Switches_7",
                           GateLockedFeedback := "F_Lock_FB_DB_7".GUARD_SWITCH.E_STOP,
                           NoEStop := "F_Lock_FB_DB_7".ESTOP.Q,
                           I_G1_GuardOpen := "Guard Position_7",
                           I_L1_Unlocked := "Lock Position_7",
                           FaultResetCmd := "Reset_Locks",
                           AllDrivesHealthy := TRUE,
                           SafetyResetDone := "F_Lock_FB_DB_7".ESTOP.Q,
                           NoVTDLocalMode := TRUE,
                           NoCrossoverPaused := TRUE,
                           Safe_Bypassed := TRUE,
                           LGX_Secure_Access := TRUE,
                           AllDevicesStopped := TRUE,
                           Gate_Station := "Control_DB".Gate_Station[7],
                           Lamps => "Lamps_7",
                           O_S1_SolenoidEnergise => "Solenoid Enable_7",
                           "Lock Reset" => "Lock Reset_7",
                           ENO => #_w1);
   "GateAccess_Station_FB_DB_8"(EN := #_w1,   // "GateAccess_Station_FB"
                           Right_True := false,
                           Switches := "Switches_8",
                           GateLockedFeedback := "F_Lock_FB_DB_8".GUARD_SWITCH.E_STOP,
                           NoEStop := "F_Lock_FB_DB_8".ESTOP.Q,
                           I_G1_GuardOpen := "Guard Position_8",
                           I_L1_Unlocked := "Lock Position_8",
                           FaultResetCmd := "Reset_Locks",
                           AllDrivesHealthy := TRUE,
                           SafetyResetDone := "F_Lock_FB_DB_8".ESTOP.Q,
                           NoVTDLocalMode := TRUE,
                           NoCrossoverPaused := TRUE,
                           Safe_Bypassed := TRUE,
                           LGX_Secure_Access := TRUE,
                           AllDevicesStopped := TRUE,
                           Gate_Station := "Control_DB".Gate_Station[8],
                           Lamps => "Lamps_8",
                           O_S1_SolenoidEnergise => "Solenoid Enable_8",
                           "Lock Reset" => "Lock Reset_8",
                           ENO => #_w2);
   "GateAccess_Station_FB_DB_11"(EN := #_w2,   // "GateAccess_Station_FB"
                           Right_True := true,
                           Switches := "Switches_11",
                           GateLockedFeedback := "F_Lock_FB_DB_11".GUARD_SWITCH.E_STOP,
                           NoEStop := "F_Lock_FB_DB_11".ESTOP.Q,
                           I_G1_GuardOpen := "Guard Position_11",
                           I_L1_Unlocked := "Lock Position_11",
                           FaultResetCmd := "Reset_Locks",
                           AllDrivesHealthy := TRUE,
                           SafetyResetDone := "F_Lock_FB_DB_11".ESTOP.Q,
                           NoVTDLocalMode := TRUE,
                           NoCrossoverPaused := TRUE,
                           Safe_Bypassed := TRUE,
                           LGX_Secure_Access := TRUE,
                           AllDevicesStopped := TRUE,
                           Gate_Station := "Control_DB".Gate_Station[11],
                           Lamps => "Lamps_11",
                           O_S1_SolenoidEnergise => "Solenoid Enable_11",
                           "Lock Reset" => "Lock Reset_11",
                           ENO => #_w3);
   IF #_w3 THEN
       "GateAccess_Station_FB_DB_12"(Right_True := true,   // "GateAccess_Station_FB"
                               Switches := "Switches_12",
                               GateLockedFeedback := "F_Lock_FB_DB_12".GUARD_SWITCH.E_STOP,
                               NoEStop := "F_Lock_FB_DB_12".ESTOP.Q,
                               I_G1_GuardOpen := "Guard Position_12",
                               I_L1_Unlocked := "Lock Position_12",
                               FaultResetCmd := "Reset_Locks",
                               AllDrivesHealthy := TRUE,
                               SafetyResetDone := "F_Lock_FB_DB_12".ESTOP.Q,
                               NoVTDLocalMode := TRUE,
                               NoCrossoverPaused := TRUE,
                               Safe_Bypassed := TRUE,
                               LGX_Secure_Access := TRUE,
                               AllDevicesStopped := TRUE,
                               Gate_Station := "Control_DB".Gate_Station[12],
                               Lamps => "Lamps_12",
                               O_S1_SolenoidEnergise => "Solenoid Enable_12",
                               "Lock Reset" => "Lock Reset_12");
   END_IF;
END_REGION

REGION Network 54: Order Tables System
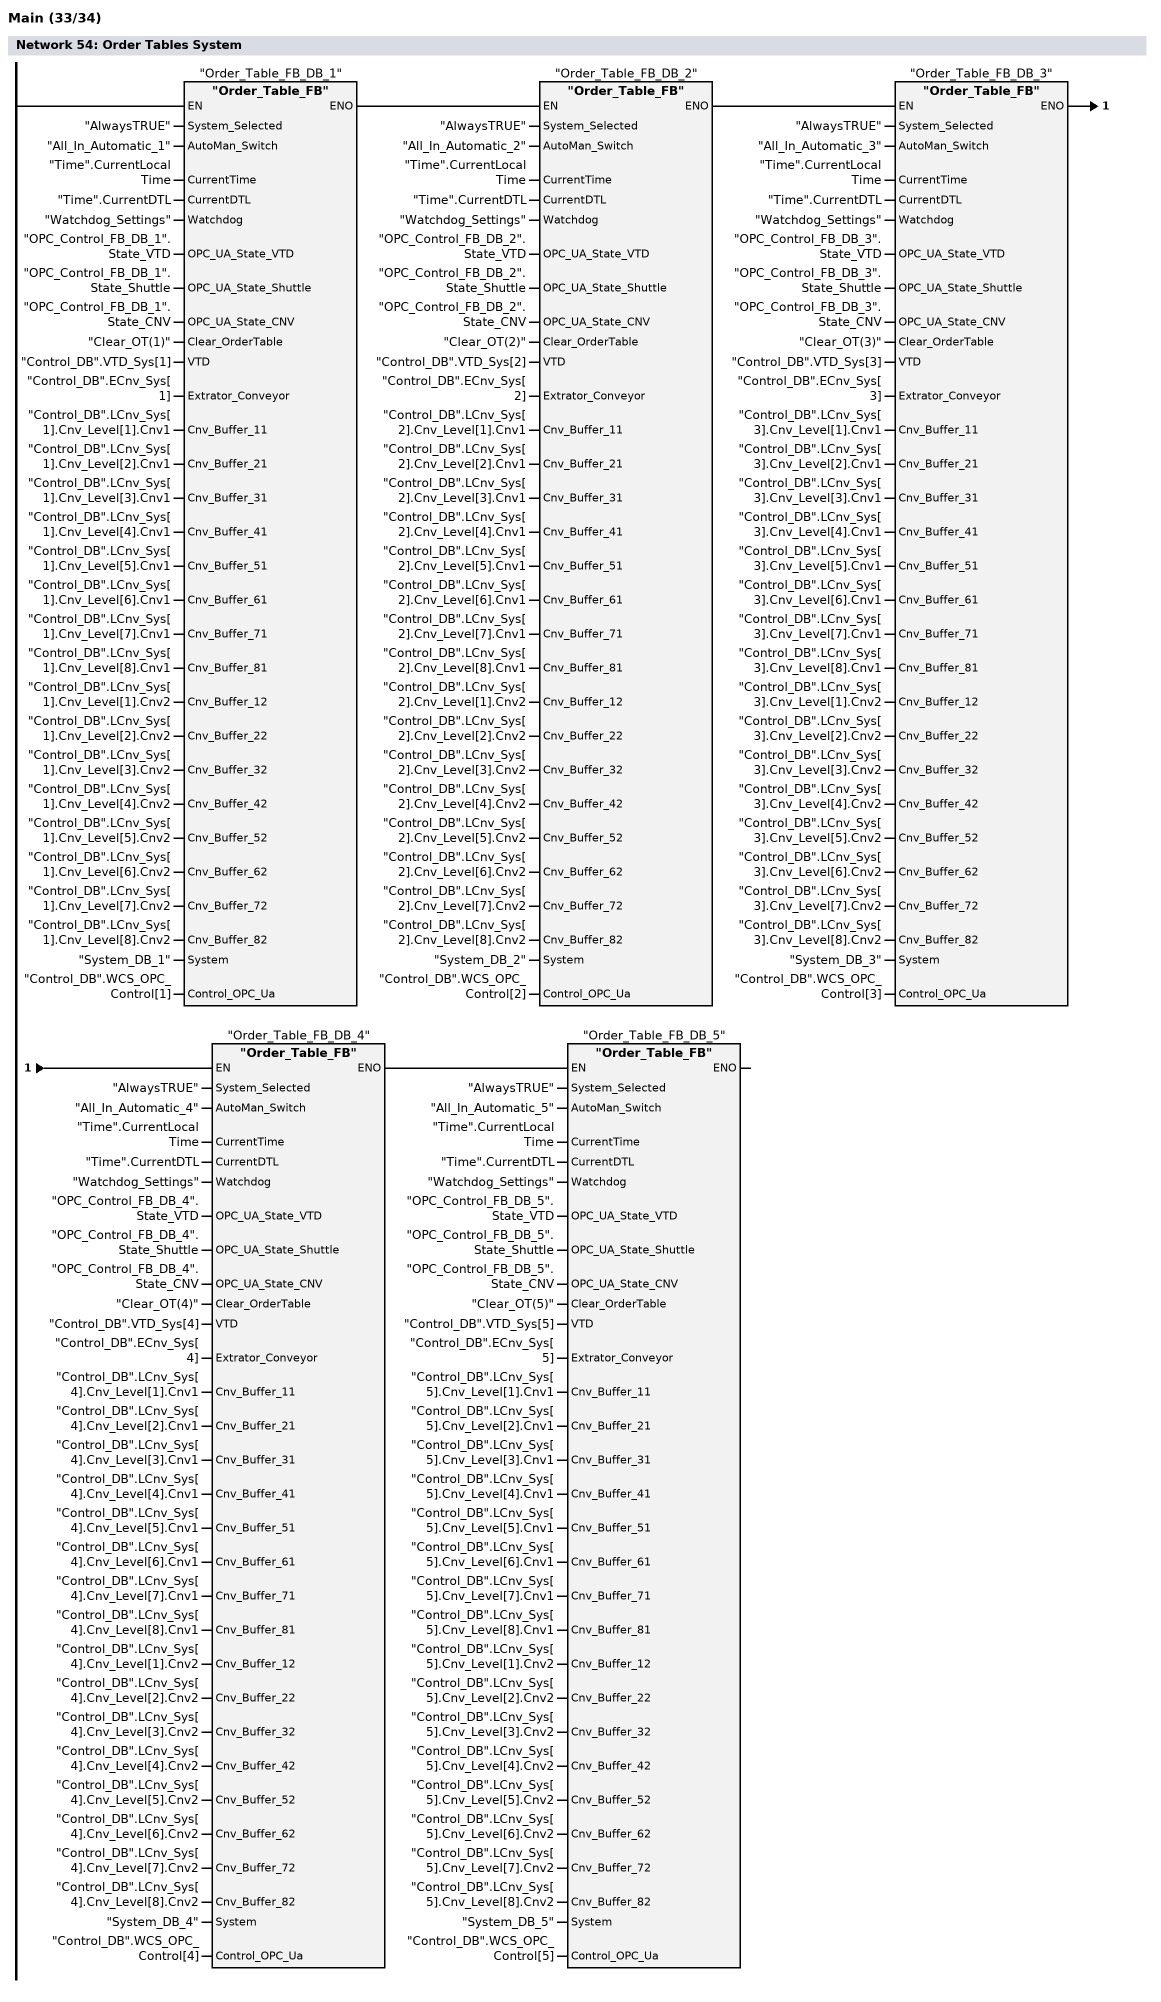
   RUNG wire#powerrail
      "Order_Table_FB_DB_1"(System_Selected := "AlwaysTRUE", AutoMan_Switch := "All_In_Automatic_1", CurrentTime := "Time".CurrentLocalTime, CurrentDTL := "Time".CurrentDTL, Watchdog := "Watchdog_Settings", OPC_UA_State_VTD := "OPC_Control_FB_DB_1".State_VTD, OPC_UA_State_Shuttle := "OPC_Control_FB_DB_1".State_Shuttle, OPC_UA_State_CNV := "OPC_Control_FB_DB_1".State_CNV, Clear_OrderTable := "Clear_OT(1)", VTD := "Control_DB".VTD_Sys[1], Extrator_Conveyor := "Control_DB".ECnv_Sys[1], Cnv_Buffer_11 := "Control_DB".LCnv_Sys[1].Cnv_Level[1].Cnv1, Cnv_Buffer_21 := "Control_DB".LCnv_Sys[1].Cnv_Level[2].Cnv1, Cnv_Buffer_31 := "Control_DB".LCnv_Sys[1].Cnv_Level[3].Cnv1, Cnv_Buffer_41 := "Control_DB".LCnv_Sys[1].Cnv_Level[4].Cnv1, Cnv_Buffer_51 := "Control_DB".LCnv_Sys[1].Cnv_Level[5].Cnv1, Cnv_Buffer_61 := "Control_DB".LCnv_Sys[1].Cnv_Level[6].Cnv1, Cnv_Buffer_71 := "Control_DB".LCnv_Sys[1].Cnv_Level[7].Cnv1, Cnv_Buffer_81 := "Control_DB".LCnv_Sys[1].Cnv_Level[8].Cnv1, Cnv_Buffer_12 := "Control_DB".LCnv_Sys[1].Cnv_Level[1].Cnv2, Cnv_Buffer_22 := "Control_DB".LCnv_Sys[1].Cnv_Level[2].Cnv2, Cnv_Buffer_32 := "Control_DB".LCnv_Sys[1].Cnv_Level[3].Cnv2, Cnv_Buffer_42 := "Control_DB".LCnv_Sys[1].Cnv_Level[4].Cnv2, Cnv_Buffer_52 := "Control_DB".LCnv_Sys[1].Cnv_Level[5].Cnv2, Cnv_Buffer_62 := "Control_DB".LCnv_Sys[1].Cnv_Level[6].Cnv2, Cnv_Buffer_72 := "Control_DB".LCnv_Sys[1].Cnv_Level[7].Cnv2, Cnv_Buffer_82 := "Control_DB".LCnv_Sys[1].Cnv_Level[8].Cnv2, System := "System_DB_1", Control_OPC_Ua := "Control_DB".WCS_OPC_Control[1])
      "Order_Table_FB_DB_2"(System_Selected := "AlwaysTRUE", AutoMan_Switch := "All_In_Automatic_2", CurrentTime := "Time".CurrentLocalTime, CurrentDTL := "Time".CurrentDTL, Watchdog := "Watchdog_Settings", OPC_UA_State_VTD := "OPC_Control_FB_DB_2".State_VTD, OPC_UA_State_Shuttle := "OPC_Control_FB_DB_2".State_Shuttle, OPC_UA_State_CNV := "OPC_Control_FB_DB_2".State_CNV, Clear_OrderTable := "Clear_OT(2)", VTD := "Control_DB".VTD_Sys[2], Extrator_Conveyor := "Control_DB".ECnv_Sys[2], Cnv_Buffer_11 := "Control_DB".LCnv_Sys[2].Cnv_Level[1].Cnv1, Cnv_Buffer_21 := "Control_DB".LCnv_Sys[2].Cnv_Level[2].Cnv1, Cnv_Buffer_31 := "Control_DB".LCnv_Sys[2].Cnv_Level[3].Cnv1, Cnv_Buffer_41 := "Control_DB".LCnv_Sys[2].Cnv_Level[4].Cnv1, Cnv_Buffer_51 := "Control_DB".LCnv_Sys[2].Cnv_Level[5].Cnv1, Cnv_Buffer_61 := "Control_DB".LCnv_Sys[2].Cnv_Level[6].Cnv1, Cnv_Buffer_71 := "Control_DB".LCnv_Sys[2].Cnv_Level[7].Cnv1, Cnv_Buffer_81 := "Control_DB".LCnv_Sys[2].Cnv_Level[8].Cnv1, Cnv_Buffer_12 := "Control_DB".LCnv_Sys[2].Cnv_Level[1].Cnv2, Cnv_Buffer_22 := "Control_DB".LCnv_Sys[2].Cnv_Level[2].Cnv2, Cnv_Buffer_32 := "Control_DB".LCnv_Sys[2].Cnv_Level[3].Cnv2, Cnv_Buffer_42 := "Control_DB".LCnv_Sys[2].Cnv_Level[4].Cnv2, Cnv_Buffer_52 := "Control_DB".LCnv_Sys[2].Cnv_Level[5].Cnv2, Cnv_Buffer_62 := "Control_DB".LCnv_Sys[2].Cnv_Level[6].Cnv2, Cnv_Buffer_72 := "Control_DB".LCnv_Sys[2].Cnv_Level[7].Cnv2, Cnv_Buffer_82 := "Control_DB".LCnv_Sys[2].Cnv_Level[8].Cnv2, System := "System_DB_2", Control_OPC_Ua := "Control_DB".WCS_OPC_Control[2])
      "Order_Table_FB_DB_3"(System_Selected := "AlwaysTRUE", AutoMan_Switch := "All_In_Automatic_3", CurrentTime := "Time".CurrentLocalTime, CurrentDTL := "Time".CurrentDTL, Watchdog := "Watchdog_Settings", OPC_UA_State_VTD := "OPC_Control_FB_DB_3".State_VTD, OPC_UA_State_Shuttle := "OPC_Control_FB_DB_3".State_Shuttle, OPC_UA_State_CNV := "OPC_Control_FB_DB_3".State_CNV, Clear_OrderTable := "Clear_OT(3)", VTD := "Control_DB".VTD_Sys[3], Extrator_Conveyor := "Control_DB".ECnv_Sys[3], Cnv_Buffer_11 := "Control_DB".LCnv_Sys[3].Cnv_Level[1].Cnv1, Cnv_Buffer_21 := "Control_DB".LCnv_Sys[3].Cnv_Level[2].Cnv1, Cnv_Buffer_31 := "Control_DB".LCnv_Sys[3].Cnv_Level[3].Cnv1, Cnv_Buffer_41 := "Control_DB".LCnv_Sys[3].Cnv_Level[4].Cnv1, Cnv_Buffer_51 := "Control_DB".LCnv_Sys[3].Cnv_Level[5].Cnv1, Cnv_Buffer_61 := "Control_DB".LCnv_Sys[3].Cnv_Level[6].Cnv1, Cnv_Buffer_71 := "Control_DB".LCnv_Sys[3].Cnv_Level[7].Cnv1, Cnv_Buffer_81 := "Control_DB".LCnv_Sys[3].Cnv_Level[8].Cnv1, Cnv_Buffer_12 := "Control_DB".LCnv_Sys[3].Cnv_Level[1].Cnv2, Cnv_Buffer_22 := "Control_DB".LCnv_Sys[3].Cnv_Level[2].Cnv2, Cnv_Buffer_32 := "Control_DB".LCnv_Sys[3].Cnv_Level[3].Cnv2, Cnv_Buffer_42 := "Control_DB".LCnv_Sys[3].Cnv_Level[4].Cnv2, Cnv_Buffer_52 := "Control_DB".LCnv_Sys[3].Cnv_Level[5].Cnv2, Cnv_Buffer_62 := "Control_DB".LCnv_Sys[3].Cnv_Level[6].Cnv2, Cnv_Buffer_72 := "Control_DB".LCnv_Sys[3].Cnv_Level[7].Cnv2, Cnv_Buffer_82 := "Control_DB".LCnv_Sys[3].Cnv_Level[8].Cnv2, System := "System_DB_3", Control_OPC_Ua := "Control_DB".WCS_OPC_Control[3])
      "Order_Table_FB_DB_4"(System_Selected := "AlwaysTRUE", AutoMan_Switch := "All_In_Automatic_4", CurrentTime := "Time".CurrentLocalTime, CurrentDTL := "Time".CurrentDTL, Watchdog := "Watchdog_Settings", OPC_UA_State_VTD := "OPC_Control_FB_DB_4".State_VTD, OPC_UA_State_Shuttle := "OPC_Control_FB_DB_4".State_Shuttle, OPC_UA_State_CNV := "OPC_Control_FB_DB_4".State_CNV, Clear_OrderTable := "Clear_OT(4)", VTD := "Control_DB".VTD_Sys[4], Extrator_Conveyor := "Control_DB".ECnv_Sys[4], Cnv_Buffer_11 := "Control_DB".LCnv_Sys[4].Cnv_Level[1].Cnv1, Cnv_Buffer_21 := "Control_DB".LCnv_Sys[4].Cnv_Level[2].Cnv1, Cnv_Buffer_31 := "Control_DB".LCnv_Sys[4].Cnv_Level[3].Cnv1, Cnv_Buffer_41 := "Control_DB".LCnv_Sys[4].Cnv_Level[4].Cnv1, Cnv_Buffer_51 := "Control_DB".LCnv_Sys[4].Cnv_Level[5].Cnv1, Cnv_Buffer_61 := "Control_DB".LCnv_Sys[4].Cnv_Level[6].Cnv1, Cnv_Buffer_71 := "Control_DB".LCnv_Sys[4].Cnv_Level[7].Cnv1, Cnv_Buffer_81 := "Control_DB".LCnv_Sys[4].Cnv_Level[8].Cnv1, Cnv_Buffer_12 := "Control_DB".LCnv_Sys[4].Cnv_Level[1].Cnv2, Cnv_Buffer_22 := "Control_DB".LCnv_Sys[4].Cnv_Level[2].Cnv2, Cnv_Buffer_32 := "Control_DB".LCnv_Sys[4].Cnv_Level[3].Cnv2, Cnv_Buffer_42 := "Control_DB".LCnv_Sys[4].Cnv_Level[4].Cnv2, Cnv_Buffer_52 := "Control_DB".LCnv_Sys[4].Cnv_Level[5].Cnv2, Cnv_Buffer_62 := "Control_DB".LCnv_Sys[4].Cnv_Level[6].Cnv2, Cnv_Buffer_72 := "Control_DB".LCnv_Sys[4].Cnv_Level[7].Cnv2, Cnv_Buffer_82 := "Control_DB".LCnv_Sys[4].Cnv_Level[8].Cnv2, System := "System_DB_4", Control_OPC_Ua := "Control_DB".WCS_OPC_Control[4])
      "Order_Table_FB_DB_5"(System_Selected := "AlwaysTRUE", AutoMan_Switch := "All_In_Automatic_5", CurrentTime := "Time".CurrentLocalTime, CurrentDTL := "Time".CurrentDTL, Watchdog := "Watchdog_Settings", OPC_UA_State_VTD := "OPC_Control_FB_DB_5".State_VTD, OPC_UA_State_Shuttle := "OPC_Control_FB_DB_5".State_Shuttle, OPC_UA_State_CNV := "OPC_Control_FB_DB_5".State_CNV, Clear_OrderTable := "Clear_OT(5)", VTD := "Control_DB".VTD_Sys[5], Extrator_Conveyor := "Control_DB".ECnv_Sys[5], Cnv_Buffer_11 := "Control_DB".LCnv_Sys[5].Cnv_Level[1].Cnv1, Cnv_Buffer_21 := "Control_DB".LCnv_Sys[5].Cnv_Level[2].Cnv1, Cnv_Buffer_31 := "Control_DB".LCnv_Sys[5].Cnv_Level[3].Cnv1, Cnv_Buffer_41 := "Control_DB".LCnv_Sys[5].Cnv_Level[4].Cnv1, Cnv_Buffer_51 := "Control_DB".LCnv_Sys[5].Cnv_Level[5].Cnv1, Cnv_Buffer_61 := "Control_DB".LCnv_Sys[5].Cnv_Level[6].Cnv1, Cnv_Buffer_71 := "Control_DB".LCnv_Sys[5].Cnv_Level[7].Cnv1, Cnv_Buffer_81 := "Control_DB".LCnv_Sys[5].Cnv_Level[8].Cnv1, Cnv_Buffer_12 := "Control_DB".LCnv_Sys[5].Cnv_Level[1].Cnv2, Cnv_Buffer_22 := "Control_DB".LCnv_Sys[5].Cnv_Level[2].Cnv2, Cnv_Buffer_32 := "Control_DB".LCnv_Sys[5].Cnv_Level[3].Cnv2, Cnv_Buffer_42 := "Control_DB".LCnv_Sys[5].Cnv_Level[4].Cnv2, Cnv_Buffer_52 := "Control_DB".LCnv_Sys[5].Cnv_Level[5].Cnv2, Cnv_Buffer_62 := "Control_DB".LCnv_Sys[5].Cnv_Level[6].Cnv2, Cnv_Buffer_72 := "Control_DB".LCnv_Sys[5].Cnv_Level[7].Cnv2, Cnv_Buffer_82 := "Control_DB".LCnv_Sys[5].Cnv_Level[8].Cnv2, System := "System_DB_5", Control_OPC_Ua := "Control_DB".WCS_OPC_Control[5])
   END_RUNG
   // the same network as SCL:
   "Order_Table_FB_DB_1"(System_Selected := "AlwaysTRUE",   // "Order_Table_FB"
                         AutoMan_Switch := "All_In_Automatic_1",
                         CurrentTime := "Time".CurrentLocalTime,
                         CurrentDTL := "Time".CurrentDTL,
                         Watchdog := "Watchdog_Settings",
                         OPC_UA_State_VTD := "OPC_Control_FB_DB_1".State_VTD,
                         OPC_UA_State_Shuttle := "OPC_Control_FB_DB_1".State_Shuttle,
                         OPC_UA_State_CNV := "OPC_Control_FB_DB_1".State_CNV,
                         Clear_OrderTable := "Clear_OT(1)",
                         VTD := "Control_DB".VTD_Sys[1],
                         Extrator_Conveyor := "Control_DB".ECnv_Sys[1],
                         Cnv_Buffer_11 := "Control_DB".LCnv_Sys[1].Cnv_Level[1].Cnv1,
                         Cnv_Buffer_21 := "Control_DB".LCnv_Sys[1].Cnv_Level[2].Cnv1,
                         Cnv_Buffer_31 := "Control_DB".LCnv_Sys[1].Cnv_Level[3].Cnv1,
                         Cnv_Buffer_41 := "Control_DB".LCnv_Sys[1].Cnv_Level[4].Cnv1,
                         Cnv_Buffer_51 := "Control_DB".LCnv_Sys[1].Cnv_Level[5].Cnv1,
                         Cnv_Buffer_61 := "Control_DB".LCnv_Sys[1].Cnv_Level[6].Cnv1,
                         Cnv_Buffer_71 := "Control_DB".LCnv_Sys[1].Cnv_Level[7].Cnv1,
                         Cnv_Buffer_81 := "Control_DB".LCnv_Sys[1].Cnv_Level[8].Cnv1,
                         Cnv_Buffer_12 := "Control_DB".LCnv_Sys[1].Cnv_Level[1].Cnv2,
                         Cnv_Buffer_22 := "Control_DB".LCnv_Sys[1].Cnv_Level[2].Cnv2,
                         Cnv_Buffer_32 := "Control_DB".LCnv_Sys[1].Cnv_Level[3].Cnv2,
                         Cnv_Buffer_42 := "Control_DB".LCnv_Sys[1].Cnv_Level[4].Cnv2,
                         Cnv_Buffer_52 := "Control_DB".LCnv_Sys[1].Cnv_Level[5].Cnv2,
                         Cnv_Buffer_62 := "Control_DB".LCnv_Sys[1].Cnv_Level[6].Cnv2,
                         Cnv_Buffer_72 := "Control_DB".LCnv_Sys[1].Cnv_Level[7].Cnv2,
                         Cnv_Buffer_82 := "Control_DB".LCnv_Sys[1].Cnv_Level[8].Cnv2,
                         System := "System_DB_1",
                         Control_OPC_Ua := "Control_DB".WCS_OPC_Control[1],
                         ENO => #_w1);
   "Order_Table_FB_DB_2"(EN := #_w1,   // "Order_Table_FB"
                         System_Selected := "AlwaysTRUE",
                         AutoMan_Switch := "All_In_Automatic_2",
                         CurrentTime := "Time".CurrentLocalTime,
                         CurrentDTL := "Time".CurrentDTL,
                         Watchdog := "Watchdog_Settings",
                         OPC_UA_State_VTD := "OPC_Control_FB_DB_2".State_VTD,
                         OPC_UA_State_Shuttle := "OPC_Control_FB_DB_2".State_Shuttle,
                         OPC_UA_State_CNV := "OPC_Control_FB_DB_2".State_CNV,
                         Clear_OrderTable := "Clear_OT(2)",
                         VTD := "Control_DB".VTD_Sys[2],
                         Extrator_Conveyor := "Control_DB".ECnv_Sys[2],
                         Cnv_Buffer_11 := "Control_DB".LCnv_Sys[2].Cnv_Level[1].Cnv1,
                         Cnv_Buffer_21 := "Control_DB".LCnv_Sys[2].Cnv_Level[2].Cnv1,
                         Cnv_Buffer_31 := "Control_DB".LCnv_Sys[2].Cnv_Level[3].Cnv1,
                         Cnv_Buffer_41 := "Control_DB".LCnv_Sys[2].Cnv_Level[4].Cnv1,
                         Cnv_Buffer_51 := "Control_DB".LCnv_Sys[2].Cnv_Level[5].Cnv1,
                         Cnv_Buffer_61 := "Control_DB".LCnv_Sys[2].Cnv_Level[6].Cnv1,
                         Cnv_Buffer_71 := "Control_DB".LCnv_Sys[2].Cnv_Level[7].Cnv1,
                         Cnv_Buffer_81 := "Control_DB".LCnv_Sys[2].Cnv_Level[8].Cnv1,
                         Cnv_Buffer_12 := "Control_DB".LCnv_Sys[2].Cnv_Level[1].Cnv2,
                         Cnv_Buffer_22 := "Control_DB".LCnv_Sys[2].Cnv_Level[2].Cnv2,
                         Cnv_Buffer_32 := "Control_DB".LCnv_Sys[2].Cnv_Level[3].Cnv2,
                         Cnv_Buffer_42 := "Control_DB".LCnv_Sys[2].Cnv_Level[4].Cnv2,
                         Cnv_Buffer_52 := "Control_DB".LCnv_Sys[2].Cnv_Level[5].Cnv2,
                         Cnv_Buffer_62 := "Control_DB".LCnv_Sys[2].Cnv_Level[6].Cnv2,
                         Cnv_Buffer_72 := "Control_DB".LCnv_Sys[2].Cnv_Level[7].Cnv2,
                         Cnv_Buffer_82 := "Control_DB".LCnv_Sys[2].Cnv_Level[8].Cnv2,
                         System := "System_DB_2",
                         Control_OPC_Ua := "Control_DB".WCS_OPC_Control[2],
                         ENO => #_w2);
   "Order_Table_FB_DB_3"(EN := #_w2,   // "Order_Table_FB"
                         System_Selected := "AlwaysTRUE",
                         AutoMan_Switch := "All_In_Automatic_3",
                         CurrentTime := "Time".CurrentLocalTime,
                         CurrentDTL := "Time".CurrentDTL,
                         Watchdog := "Watchdog_Settings",
                         OPC_UA_State_VTD := "OPC_Control_FB_DB_3".State_VTD,
                         OPC_UA_State_Shuttle := "OPC_Control_FB_DB_3".State_Shuttle,
                         OPC_UA_State_CNV := "OPC_Control_FB_DB_3".State_CNV,
                         Clear_OrderTable := "Clear_OT(3)",
                         VTD := "Control_DB".VTD_Sys[3],
                         Extrator_Conveyor := "Control_DB".ECnv_Sys[3],
                         Cnv_Buffer_11 := "Control_DB".LCnv_Sys[3].Cnv_Level[1].Cnv1,
                         Cnv_Buffer_21 := "Control_DB".LCnv_Sys[3].Cnv_Level[2].Cnv1,
                         Cnv_Buffer_31 := "Control_DB".LCnv_Sys[3].Cnv_Level[3].Cnv1,
                         Cnv_Buffer_41 := "Control_DB".LCnv_Sys[3].Cnv_Level[4].Cnv1,
                         Cnv_Buffer_51 := "Control_DB".LCnv_Sys[3].Cnv_Level[5].Cnv1,
                         Cnv_Buffer_61 := "Control_DB".LCnv_Sys[3].Cnv_Level[6].Cnv1,
                         Cnv_Buffer_71 := "Control_DB".LCnv_Sys[3].Cnv_Level[7].Cnv1,
                         Cnv_Buffer_81 := "Control_DB".LCnv_Sys[3].Cnv_Level[8].Cnv1,
                         Cnv_Buffer_12 := "Control_DB".LCnv_Sys[3].Cnv_Level[1].Cnv2,
                         Cnv_Buffer_22 := "Control_DB".LCnv_Sys[3].Cnv_Level[2].Cnv2,
                         Cnv_Buffer_32 := "Control_DB".LCnv_Sys[3].Cnv_Level[3].Cnv2,
                         Cnv_Buffer_42 := "Control_DB".LCnv_Sys[3].Cnv_Level[4].Cnv2,
                         Cnv_Buffer_52 := "Control_DB".LCnv_Sys[3].Cnv_Level[5].Cnv2,
                         Cnv_Buffer_62 := "Control_DB".LCnv_Sys[3].Cnv_Level[6].Cnv2,
                         Cnv_Buffer_72 := "Control_DB".LCnv_Sys[3].Cnv_Level[7].Cnv2,
                         Cnv_Buffer_82 := "Control_DB".LCnv_Sys[3].Cnv_Level[8].Cnv2,
                         System := "System_DB_3",
                         Control_OPC_Ua := "Control_DB".WCS_OPC_Control[3],
                         ENO => #_w3);
   "Order_Table_FB_DB_4"(EN := #_w3,   // "Order_Table_FB"
                         System_Selected := "AlwaysTRUE",
                         AutoMan_Switch := "All_In_Automatic_4",
                         CurrentTime := "Time".CurrentLocalTime,
                         CurrentDTL := "Time".CurrentDTL,
                         Watchdog := "Watchdog_Settings",
                         OPC_UA_State_VTD := "OPC_Control_FB_DB_4".State_VTD,
                         OPC_UA_State_Shuttle := "OPC_Control_FB_DB_4".State_Shuttle,
                         OPC_UA_State_CNV := "OPC_Control_FB_DB_4".State_CNV,
                         Clear_OrderTable := "Clear_OT(4)",
                         VTD := "Control_DB".VTD_Sys[4],
                         Extrator_Conveyor := "Control_DB".ECnv_Sys[4],
                         Cnv_Buffer_11 := "Control_DB".LCnv_Sys[4].Cnv_Level[1].Cnv1,
                         Cnv_Buffer_21 := "Control_DB".LCnv_Sys[4].Cnv_Level[2].Cnv1,
                         Cnv_Buffer_31 := "Control_DB".LCnv_Sys[4].Cnv_Level[3].Cnv1,
                         Cnv_Buffer_41 := "Control_DB".LCnv_Sys[4].Cnv_Level[4].Cnv1,
                         Cnv_Buffer_51 := "Control_DB".LCnv_Sys[4].Cnv_Level[5].Cnv1,
                         Cnv_Buffer_61 := "Control_DB".LCnv_Sys[4].Cnv_Level[6].Cnv1,
                         Cnv_Buffer_71 := "Control_DB".LCnv_Sys[4].Cnv_Level[7].Cnv1,
                         Cnv_Buffer_81 := "Control_DB".LCnv_Sys[4].Cnv_Level[8].Cnv1,
                         Cnv_Buffer_12 := "Control_DB".LCnv_Sys[4].Cnv_Level[1].Cnv2,
                         Cnv_Buffer_22 := "Control_DB".LCnv_Sys[4].Cnv_Level[2].Cnv2,
                         Cnv_Buffer_32 := "Control_DB".LCnv_Sys[4].Cnv_Level[3].Cnv2,
                         Cnv_Buffer_42 := "Control_DB".LCnv_Sys[4].Cnv_Level[4].Cnv2,
                         Cnv_Buffer_52 := "Control_DB".LCnv_Sys[4].Cnv_Level[5].Cnv2,
                         Cnv_Buffer_62 := "Control_DB".LCnv_Sys[4].Cnv_Level[6].Cnv2,
                         Cnv_Buffer_72 := "Control_DB".LCnv_Sys[4].Cnv_Level[7].Cnv2,
                         Cnv_Buffer_82 := "Control_DB".LCnv_Sys[4].Cnv_Level[8].Cnv2,
                         System := "System_DB_4",
                         Control_OPC_Ua := "Control_DB".WCS_OPC_Control[4],
                         ENO => #_w4);
   IF #_w4 THEN
       "Order_Table_FB_DB_5"(System_Selected := "AlwaysTRUE",   // "Order_Table_FB"
                             AutoMan_Switch := "All_In_Automatic_5",
                             CurrentTime := "Time".CurrentLocalTime,
                             CurrentDTL := "Time".CurrentDTL,
                             Watchdog := "Watchdog_Settings",
                             OPC_UA_State_VTD := "OPC_Control_FB_DB_5".State_VTD,
                             OPC_UA_State_Shuttle := "OPC_Control_FB_DB_5".State_Shuttle,
                             OPC_UA_State_CNV := "OPC_Control_FB_DB_5".State_CNV,
                             Clear_OrderTable := "Clear_OT(5)",
                             VTD := "Control_DB".VTD_Sys[5],
                             Extrator_Conveyor := "Control_DB".ECnv_Sys[5],
                             Cnv_Buffer_11 := "Control_DB".LCnv_Sys[5].Cnv_Level[1].Cnv1,
                             Cnv_Buffer_21 := "Control_DB".LCnv_Sys[5].Cnv_Level[2].Cnv1,
                             Cnv_Buffer_31 := "Control_DB".LCnv_Sys[5].Cnv_Level[3].Cnv1,
                             Cnv_Buffer_41 := "Control_DB".LCnv_Sys[5].Cnv_Level[4].Cnv1,
                             Cnv_Buffer_51 := "Control_DB".LCnv_Sys[5].Cnv_Level[5].Cnv1,
                             Cnv_Buffer_61 := "Control_DB".LCnv_Sys[5].Cnv_Level[6].Cnv1,
                             Cnv_Buffer_71 := "Control_DB".LCnv_Sys[5].Cnv_Level[7].Cnv1,
                             Cnv_Buffer_81 := "Control_DB".LCnv_Sys[5].Cnv_Level[8].Cnv1,
                             Cnv_Buffer_12 := "Control_DB".LCnv_Sys[5].Cnv_Level[1].Cnv2,
                             Cnv_Buffer_22 := "Control_DB".LCnv_Sys[5].Cnv_Level[2].Cnv2,
                             Cnv_Buffer_32 := "Control_DB".LCnv_Sys[5].Cnv_Level[3].Cnv2,
                             Cnv_Buffer_42 := "Control_DB".LCnv_Sys[5].Cnv_Level[4].Cnv2,
                             Cnv_Buffer_52 := "Control_DB".LCnv_Sys[5].Cnv_Level[5].Cnv2,
                             Cnv_Buffer_62 := "Control_DB".LCnv_Sys[5].Cnv_Level[6].Cnv2,
                             Cnv_Buffer_72 := "Control_DB".LCnv_Sys[5].Cnv_Level[7].Cnv2,
                             Cnv_Buffer_82 := "Control_DB".LCnv_Sys[5].Cnv_Level[8].Cnv2,
                             System := "System_DB_5",
                             Control_OPC_Ua := "Control_DB".WCS_OPC_Control[5]);
   END_IF;
END_REGION

REGION Network 55: LOGISTEX
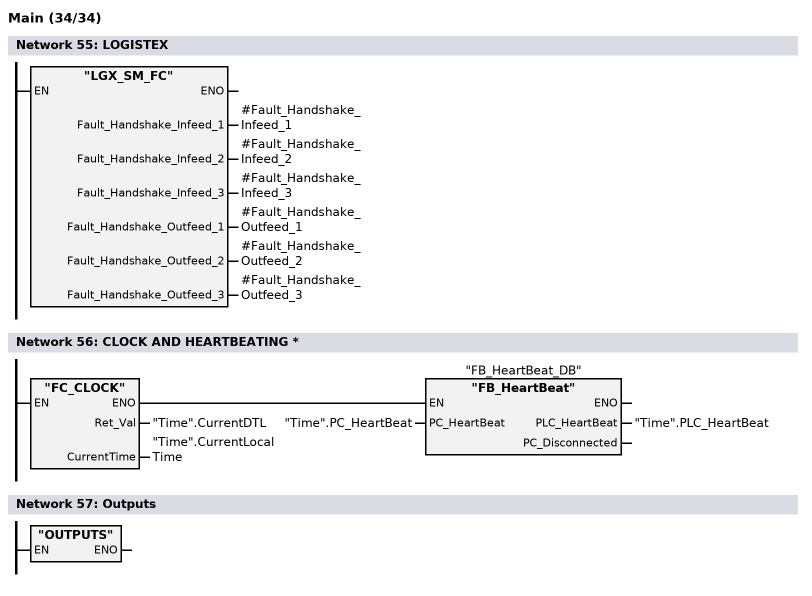
   RUNG wire#powerrail
      "LGX_SM_FC"(Fault_Handshake_Infeed_1 => #Fault_Handshake_Infeed_1, Fault_Handshake_Infeed_2 => #Fault_Handshake_Infeed_2, Fault_Handshake_Infeed_3 => #Fault_Handshake_Infeed_3, Fault_Handshake_Outfeed_1 => #Fault_Handshake_Outfeed_1, Fault_Handshake_Outfeed_2 => #Fault_Handshake_Outfeed_2, Fault_Handshake_Outfeed_3 => #Fault_Handshake_Outfeed_3)
   END_RUNG
   // the same network as SCL:
   "LGX_SM_FC"(Fault_Handshake_Infeed_1 => #Fault_Handshake_Infeed_1,
               Fault_Handshake_Infeed_2 => #Fault_Handshake_Infeed_2,
               Fault_Handshake_Infeed_3 => #Fault_Handshake_Infeed_3,
               Fault_Handshake_Outfeed_1 => #Fault_Handshake_Outfeed_1,
               Fault_Handshake_Outfeed_2 => #Fault_Handshake_Outfeed_2,
               Fault_Handshake_Outfeed_3 => #Fault_Handshake_Outfeed_3);
END_REGION

REGION Network 56: CLOCK AND HEARTBEATING *
   RUNG wire#powerrail
      "FC_CLOCK"(Ret_Val => "Time".CurrentDTL, CurrentTime => "Time".CurrentLocalTime)
      "FB_HeartBeat_DB"(PC_HeartBeat := "Time".PC_HeartBeat, PLC_HeartBeat => "Time".PLC_HeartBeat, PC_Disconnected =>)
   END_RUNG
   // the same network as SCL:
   "Time".CurrentDTL := "FC_CLOCK"(CurrentTime => "Time".CurrentLocalTime, ENO => #_w1);
   IF #_w1 THEN
       "FB_HeartBeat_DB"(PC_HeartBeat := "Time".PC_HeartBeat, PLC_HeartBeat => "Time".PLC_HeartBeat);   // "FB_HeartBeat"
   END_IF;
END_REGION

REGION Network 57: Outputs
   RUNG wire#powerrail
      "OUTPUTS"()
   END_RUNG
   // the same network as SCL:
   "OUTPUTS"();
END_REGION
END_ORGANIZATION_BLOCK

FUNCTION "INPUTS" : Void   // FC25, SCL
{ S7_Optimized_Access := 'TRUE' }
VERSION : 0.1
// stored: AutoNumber true, IsIECCheckEnabled false, SetENOAutomatically false, UDAEnableTagReadback false
BEGIN
   REGION SYSTEM 1
       REGION EXTRACTOR CONVEYOR
           "Control_DB".ECnv_Sys[1].Inputs.Left := "CVTD1 SENSOR CONVEYOR LEFT";
           "Control_DB".ECnv_Sys[1].Inputs.Lpd1 := "CVTD1 SENSOR CONVEYOR LEFT (PALLET DETECT 1)";
           "Control_DB".ECnv_Sys[1].Inputs.Center := "CVTD1 SENSOR CONVEYOR CENTER";
           "Control_DB".ECnv_Sys[1].Inputs.Right := "CVTD1 SENSOR CONVEYOR RIGHT";
           "Control_DB".ECnv_Sys[1].Inputs.Rpd1 := "CVTD1 SENSOR CONVEYOR RIGHT (PALLET DETECT 1)";

           "T_OH_Left_1".TOF(IN := "CVTD1 OVERHANG LEFT" OR NOT "Control_DB".VTD_Sys[1].Running,
                             PT := T#200ms);
           "Control_DB".ECnv_Sys[1].Inputs.Overhang_Left := "T_OH_Left_1".Q;

           "T_OH_Right_1".TOF(IN := "CVTD1 OVERHANG RIGHT" OR NOT "Control_DB".VTD_Sys[1].Running,
                              PT := T#200ms);
           "Control_DB".ECnv_Sys[1].Inputs.Overhang_Right := "T_OH_Right_1".Q;

           "Control_DB".ECnv_Sys[1].Inputs.VFD_Status := "CVTD1_StatusWord";
           "Control_DB".ECnv_Sys[1].Inputs.VFD_ActualCurrent := WORD_TO_INT("CVTD1_ActualCurrent");
           "Control_DB".ECnv_Sys[1].Inputs.VFD_Speed_Actual := WORD_TO_INT("CVTD1_ActualSpeed");
           "Control_DB".ECnv_Sys[1].Inputs.VFD_ActualTorque := WORD_TO_INT("CVTD1_ActualTorque");
       END_REGION

